(* IEC 61131-3 sources: Industry-PLC-LLM/data/PLCBEAD_repo/PLCBEAD_PLCEmbed-main/PLC-BEAD/Source/PLC_Programs (part 2) *)

(* ---- ALARM_2.ST ---- *)
FUNCTION_BLOCK ALARM_2
	VAR_INPUT
		X :	REAL;
		LO_1 :	REAL;
		HI_1 :	REAL;
		LO_2 :	REAL;
		HI_2 :	REAL;
		HYS :	REAL;
	END_VAR

	VAR_OUTPUT
		Q1_LO :	BOOL;
		Q1_HI :	BOOL;
		Q2_LO :	BOOL;
		Q2_HI :	BOOL;
	END_VAR

	VAR
		tmp :	REAL;
	END_VAR

	tmp := X - Hys * 0.5;
	IF tmp > LO_1 THEN Q1_LO := FALSE; END_IF;
	IF tmp > LO_2 THEN Q2_LO := FALSE; END_IF;
	IF tmp > HI_1 THEN Q1_HI := TRUE; END_IF;
	IF tmp > HI_2 THEN Q2_HI := TRUE; END_IF;
	tmp := tmp + hys;
	IF tmp < LO_1 THEN Q1_LO := TRUE; END_IF;
	IF tmp < LO_2 THEN Q2_LO := TRUE; END_IF;
	IF tmp < HI_1 THEN Q1_HI := FALSE; END_IF;
	IF tmp < HI_2 THEN Q2_HI := FALSE; END_IF;

END_FUNCTION_BLOCK

PROGRAM program0
	VAR
	    LocalVar0 : REAL;
		LocalVar1 : REAL;
		LocalVar2 : REAL;
		LocalVar3 : REAL;
		LocalVar4 : REAL;
		LocalVar5 : REAL;
		LocalOUT1  : BOOL;
		LocalOUT2  : BOOL;
		LocalOUT3  : BOOL;
		LocalOUT4  : BOOL;
		func_block : ALARM_2;
  	END_VAR
	func_block.X := LocalVar0;
	func_block.LO_1 := LocalVar1;
	func_block.HI_1 := LocalVar2;
	func_block.LO_2 := LocalVar3;
	func_block.HI_2 := LocalVar4;
	func_block.HYS := LocalVar5;
	func_block();
	LocalOUT1 := func_block.Q1_LO;
	LocalOUT2 := func_block.Q1_HI;
	LocalOUT3 := func_block.Q2_LO;
	LocalOUT4 := func_block.Q2_HI;
END_PROGRAM

CONFIGURATION Config0
  	RESOURCE Res0 ON PLC
    	TASK task0(INTERVAL := T#20ms,PRIORITY := 0);
    	PROGRAM instance0 WITH task0 : program0;
  	END_RESOURCE
END_CONFIGURATION

(* ---- ARRAY_AVG.ST ---- *)
TYPE
	oscat_pt_ARRAY: ARRAY [1..100] OF REAL;
END_TYPE

FUNCTION_BLOCK ARRAY_AVG_Block
	VAR_IN_OUT
		PT :	oscat_pt_ARRAY;
	END_VAR

	VAR_INPUT
		SIZE :	UINT;
	END_VAR

	VAR_OUTPUT
		ARRAY_AVG :	REAL;
	END_VAR

	VAR
		i :	INT;
		stop :	INT;
	END_VAR

	stop :=LIMIT_INT(1,UINT_TO_INT(size),1000);

	array_avg := 0.0;
	FOR i := 1 TO stop DO
		array_avg := array_avg + pt[i];
	END_FOR;
	array_avg := array_avg / INT_TO_REAL(stop);
END_FUNCTION_BLOCK

PROGRAM program0
  VAR
    LocalVar0 : oscat_pt_ARRAY;
    LocalVar1 : UINT;
	LocalOUT  : REAL;
	func_block : ARRAY_AVG_Block;
  END_VAR
	func_block.pt := LocalVar0;
	func_block.size := LocalVar1;
	func_block();
	LocalOUT := func_block.ARRAY_AVG;

END_PROGRAM

CONFIGURATION Config0
  RESOURCE Res0 ON PLC
    TASK task0(INTERVAL := T#20ms,PRIORITY := 0);
    PROGRAM instance0 WITH task0 : program0;
  END_RESOURCE
END_CONFIGURATION

(* ---- ARRAY_GAV.ST ---- *)
TYPE
	oscat_pt_ARRAY: ARRAY [1..100] OF REAL;
END_TYPE

FUNCTION SQRTN:REAL
	VAR_INPUT
		X :	REAL;
		N :	INT;
	END_VAR

	IF N > 0 THEN
		SQRTN := EXP(LN(x) / INT_TO_REAL(n));
	ELSE
		SQRTN := 0.0;
	END_IF;
END_FUNCTION

FUNCTION_BLOCK ARRAY_GAV_Block
	VAR_IN_OUT
		PT :	oscat_pt_ARRAY;
	END_VAR

	VAR_INPUT
		SIZE :	UINT;
	END_VAR

	VAR_OUTPUT
		ARRAY_GAV :	REAL;
	END_VAR

	VAR
		i :	INT;
		stop :	INT;
	END_VAR

	stop :=LIMIT_INT(1,UINT_TO_INT(size),1000);
	ARRAY_GAV := 1.0;
	FOR i := 1 TO stop DO
		IF pt[i] > 0.0 THEN
			ARRAY_GAV := ARRAY_GAV * pt[i];
		ELSE
			ARRAY_GAV := 0.0;
			RETURN;
		END_IF;
	END_FOR;
	ARRAY_GAV := SQRTN(ARRAY_GAV,stop);
END_FUNCTION_BLOCK

PROGRAM program0
  VAR
    LocalVar0 : oscat_pt_ARRAY;
    LocalVar1 : UINT;
	LocalOUT  : REAL;
	func_block : ARRAY_GAV_Block;
  END_VAR
	func_block.pt := LocalVar0;
	func_block.size := LocalVar1;
	func_block();
	LocalOUT := func_block.ARRAY_GAV;

END_PROGRAM

CONFIGURATION Config0
  RESOURCE Res0 ON PLC
    TASK task0(INTERVAL := T#20ms,PRIORITY := 0);
    PROGRAM instance0 WITH task0 : program0;
  END_RESOURCE
END_CONFIGURATION

(* ---- ARRAY_HAV.ST ---- *)
TYPE
	oscat_pt_ARRAY: ARRAY [1..100] OF REAL;
END_TYPE

FUNCTION_BLOCK ARRAY_HAV_Block
	VAR_IN_OUT
		PT :	oscat_pt_ARRAY;
	END_VAR

	VAR_INPUT
		SIZE :	UINT;
	END_VAR

	VAR_OUTPUT
		ARRAY_HAV :	REAL;
	END_VAR

	VAR
		i :	INT;
		stop :	INT;
	END_VAR

	stop :=LIMIT_INT(1,UINT_TO_INT(size),1000);
	ARRAY_HAV := 0.0;
	FOR i := 1 TO stop DO
		IF pt[i] <> 0.0 THEN
			ARRAY_HAV := ARRAY_HAV + 1.0/pt[i];
		ELSE
			ARRAY_HAV := 0.0;
			RETURN;
		END_IF;
	END_FOR;
	ARRAY_HAV := INT_TO_REAL(stop) / ARRAY_HAV;
END_FUNCTION_BLOCK

PROGRAM program0
  VAR
    LocalVar0 : oscat_pt_ARRAY;
    LocalVar1 : UINT;
	LocalOUT  : REAL;
	func_block : ARRAY_HAV_Block;
  END_VAR
	func_block.pt := LocalVar0;
	func_block.size := LocalVar1;
	func_block();
	LocalOUT := func_block.ARRAY_HAV;

END_PROGRAM

CONFIGURATION Config0
  RESOURCE Res0 ON PLC
    TASK task0(INTERVAL := T#20ms,PRIORITY := 0);
    PROGRAM instance0 WITH task0 : program0;
  END_RESOURCE
END_CONFIGURATION

(* ---- ARRAY_MAX.ST ---- *)
TYPE
	oscat_pt_ARRAY: ARRAY [1..100] OF REAL;
END_TYPE

FUNCTION_BLOCK ARRAY_MAX_Block
	VAR_IN_OUT
		PT :	oscat_pt_ARRAY;
	END_VAR

	VAR_INPUT
		SIZE :	UINT;
	END_VAR

	VAR_OUTPUT
		ARRAY_MAX :	REAL;
	END_VAR

	VAR
		i :	INT;
		stop :	INT;
	END_VAR

	stop :=LIMIT_INT(1,UINT_TO_INT(size),1000);

	FOR i := 1 TO stop DO
		IF pt[i] > array_max THEN array_max := pt[i]; END_IF;
	END_FOR;

END_FUNCTION_BLOCK

PROGRAM program0
  VAR
    LocalVar0 : oscat_pt_ARRAY;
    LocalVar1 : UINT;
	LocalOUT  : REAL;
	func_block : ARRAY_MAX_Block;
  END_VAR
	func_block.pt := LocalVar0;
	func_block.size := LocalVar1;
	func_block();
	LocalOUT := func_block.ARRAY_MAX;

END_PROGRAM

CONFIGURATION Config0
  RESOURCE Res0 ON PLC
    TASK task0(INTERVAL := T#20ms,PRIORITY := 0);
    PROGRAM instance0 WITH task0 : program0;
  END_RESOURCE
END_CONFIGURATION

(* ---- ARRAY_MEDIAN.ST ---- *)
TYPE
	oscat_pt_ARRAY: ARRAY [1..100] OF REAL;
	oscat_stack_array: ARRAY [1..32]   OF INT;
END_TYPE

FUNCTION _INT_TO_UDINT:UDINT
	VAR_INPUT
		IN :	INT;
	END_VAR

	_INT_TO_UDINT := DINT_TO_UDINT(INT_TO_DINT(IN));
END_FUNCTION

FUNCTION BIT_OF_DWORD:BOOL
	VAR_INPUT
		IN :	DWORD;
		N :	INT;
	END_VAR
	BIT_OF_DWORD := (SHR(in,n) AND DWORD#1) > DWORD#0;
END_FUNCTION

FUNCTION EVEN:BOOL
	VAR_INPUT
		IN :	DINT;
	END_VAR
	even := NOT BIT_OF_DWORD(DINT_TO_DWORD(in),0);
END_FUNCTION

FUNCTION_BLOCK _ARRAY_SORT_Block
	VAR_IN_OUT
		PT :	oscat_pt_ARRAY;
	END_VAR

	VAR_INPUT
		SIZE :	UINT;
	END_VAR

	VAR_OUTPUT
		_ARRAY_SORT :BOOL;
	END_VAR

	VAR
		stack_count :	INT;
		stack :	oscat_stack_array;
		links :	INT;
		rechts :	INT;
		pivot :	REAL;
		i :	INT;
		j :	INT;
		ende_innen :	BOOL;
		ende_aussen :	BOOL;
		tmp :	REAL;
		x :	INT;
	END_VAR

	links := 1;
	rechts := DWORD_TO_INT(SHR(UINT_TO_DWORD(size),2));
	stack_count := 1;

	WHILE NOT ende_aussen DO
		IF links < rechts THEN
			x := DWORD_TO_INT(SHR(UDINT_TO_DWORD(_INT_TO_UDINT(rechts)+ _INT_TO_UDINT(links)),1));
			pivot := PT[x];
			i := links - 1;
			j := rechts + 1;

			ende_innen := FALSE;
			REPEAT
				REPEAT	i := i+1;	UNTIL (PT[i] >= pivot) OR NOT (i < rechts)	END_REPEAT;
				REPEAT	j := j-1;	UNTIL (PT[j] <= pivot) OR NOT (j > links)	END_REPEAT;
				IF i >= j THEN
					ende_innen := TRUE;
				ELSE
					tmp := PT[j];
					PT[j] := PT[i];
					PT[i] := tmp;
				END_IF;

			UNTIL ende_innen END_REPEAT;

			stack[stack_count] := rechts;
			IF Stack_count < 32 THEN
				stack_count := stack_count +1;
			ELSE
				ende_aussen := TRUE;
				_ARRAY_SORT := FALSE;
			END_IF;
			rechts := MAX(links, i-1);

		ELSE
			IF stack_count = 1 THEN
				ende_aussen := TRUE;
			ELSE
				links := rechts+1;
				stack_count := stack_count - 1;
				rechts:= stack[stack_count];
			END_IF;
		END_IF;
	END_WHILE;

	_ARRAY_SORT := TRUE;
END_FUNCTION_BLOCK

FUNCTION_BLOCK _ARRAY_MEDIAN_Block

	VAR_IN_OUT
		PT :	oscat_pt_ARRAY;
	END_VAR

	VAR_INPUT
		SIZE :	UINT;
	END_VAR

	VAR_OUTPUT
		_ARRAY_MEDIAN :	REAL;
	END_VAR

	VAR
		i :	INT;
		i2 :	INT;
		stop :	INT;
		_array_sort :	_ARRAY_SORT_Block;
	END_VAR

	(* Array sortieren *)
	_array_sort.pt   := pt;
	_array_sort.size := size;
	_array_sort();
	pt := _array_sort.pt;

	stop :=LIMIT_INT(1,UINT_TO_INT(size),1000);
	IF even(INT_TO_DINT(stop)) THEN
	    i := WORD_TO_INT(SHR(INT_TO_WORD(stop),1));
	    i2 := i+1;
		_array_median := (pt[i] + pt[i2]) * 0.5;
	ELSE
	    i := WORD_TO_INT(SHR(INT_TO_WORD(stop),1))+1;
		_array_median := pt[i];
	END_IF;

END_FUNCTION_BLOCK

PROGRAM program0
  VAR
    LocalVar0 : oscat_pt_ARRAY;
    LocalVar1 : UINT;
	LocalOUT  : REAL;
	func_block : _ARRAY_MEDIAN_Block;
  END_VAR
	func_block.pt := LocalVar0;
	func_block.size := LocalVar1;
	func_block();
	LocalOUT := func_block._ARRAY_MEDIAN;
	LocalVar0 := func_block.pt;

END_PROGRAM

CONFIGURATION Config0
  RESOURCE Res0 ON PLC
    TASK task0(INTERVAL := T#20ms,PRIORITY := 0);
    PROGRAM instance0 WITH task0 : program0;
  END_RESOURCE
END_CONFIGURATION

(* ---- ARRAY_MIN.ST ---- *)
TYPE
	oscat_pt_ARRAY: ARRAY [1..100] OF REAL;
END_TYPE

FUNCTION_BLOCK ARRAY_MIN_Block
	VAR_IN_OUT
		PT :	oscat_pt_ARRAY;
	END_VAR

	VAR_INPUT
		SIZE :	UINT;
	END_VAR

	VAR_OUTPUT
		ARRAY_MIN :	REAL;
	END_VAR

	VAR
		i :	INT;
		stop :	INT;
	END_VAR

	stop :=LIMIT_INT(1,UINT_TO_INT(size),1000);

	array_min := pt[1];
	FOR i := 2 TO stop DO
		IF pt[i] < array_min THEN array_min := pt[i]; END_IF;
	END_FOR;

END_FUNCTION_BLOCK
PROGRAM program0
  VAR
    LocalVar0 : oscat_pt_ARRAY;
    LocalVar1 : UINT;
	LocalOUT  : REAL;
	func_block : ARRAY_MIN_Block;
  END_VAR
	func_block.pt := LocalVar0;
	func_block.size := LocalVar1;
	func_block();
	LocalOUT := func_block.ARRAY_MIN;

END_PROGRAM

CONFIGURATION Config0
  RESOURCE Res0 ON PLC
    TASK task0(INTERVAL := T#20ms,PRIORITY := 0);
    PROGRAM instance0 WITH task0 : program0;
  END_RESOURCE
END_CONFIGURATION

(* ---- ARRAY_SDV.ST ---- *)
TYPE
	oscat_pt_ARRAY: ARRAY [1..100] OF REAL;
END_TYPE

FUNCTION_BLOCK ARRAY_VAR_Block
	VAR_IN_OUT
		PT :	oscat_pt_ARRAY;
	END_VAR

	VAR_INPUT
		SIZE :	UINT;
	END_VAR

	VAR_OUTPUT
		ARRAY_VAR :	REAL;
	END_VAR

	VAR
		i :	INT;
		stop :	INT;
		avg :	REAL;
	END_VAR

	stop :=LIMIT_INT(1,UINT_TO_INT(size),1000);
	avg := pt[1];
	FOR i := 2 TO stop DO
		avg := avg + pt[i];
	END_FOR;
	avg := avg / INT_TO_REAL(stop);

	array_var := EXPT(pt[1] - avg, 2.0);
	FOR i := 2 TO stop DO
		array_var := array_var + EXPT(pt[i] - avg, 2.0);
	END_FOR;
	array_var := array_var / INT_TO_REAL(stop-1);

END_FUNCTION_BLOCK

FUNCTION_BLOCK ARRAY_SDV_Block
	VAR_IN_OUT
		PT :	oscat_pt_ARRAY;
	END_VAR

	VAR_INPUT
		SIZE :	UINT;
	END_VAR

	VAR_OUTPUT
		ARRAY_SDV :	REAL;
	END_VAR

	VAR
		FB_array_var :	array_var_block;
	END_VAR

	FB_array_var.pt   := pt;
	FB_array_var.size := size;
	FB_array_var();
	pt := FB_array_var.pt;

	array_sdv := SQRT(FB_array_var.array_var);
END_FUNCTION_BLOCK

PROGRAM program0
  VAR
    LocalVar0 : oscat_pt_ARRAY;
    LocalVar1 : UINT;
	LocalOUT  : REAL;
	func_block : ARRAY_SDV_Block;
  END_VAR
	func_block.pt := LocalVar0;
	func_block.size := LocalVar1;
	func_block();
	LocalOUT := func_block.ARRAY_SDV;

END_PROGRAM

CONFIGURATION Config0
  RESOURCE Res0 ON PLC
    TASK task0(INTERVAL := T#20ms,PRIORITY := 0);
    PROGRAM instance0 WITH task0 : program0;
  END_RESOURCE
END_CONFIGURATION

(* ---- ARRAY_SPR.ST ---- *)
TYPE
	oscat_pt_ARRAY: ARRAY [1..100] OF REAL;
END_TYPE

FUNCTION_BLOCK ARRAY_SPR_Block
	VAR_IN_OUT
		PT :	oscat_pt_ARRAY;
	END_VAR

	VAR_INPUT
		SIZE :	UINT;
	END_VAR

	VAR_OUTPUT
		ARRAY_SPR :	REAL;
	END_VAR

	VAR
		i :	INT;
		stop :	INT;
		array_max :	REAL;
		array_min :	REAL;
	END_VAR

	stop :=LIMIT_INT(1,UINT_TO_INT(size),1000);

	array_min := pt[1];
	array_max := pt[1];
	FOR i := 2 TO stop DO
		IF pt[i] > array_max THEN array_max := pt[i];
		ELSIF pt[i] < array_min THEN array_min := pt[i];
		END_IF;
	END_FOR;
	array_spr := array_max - array_min;
END_FUNCTION_BLOCK

PROGRAM program0
  VAR
    LocalVar0 : oscat_pt_ARRAY;
    LocalVar1 : UINT;
	LocalOUT  : REAL;
	func_block : ARRAY_SPR_Block;
  END_VAR
	func_block.pt := LocalVar0;
	func_block.size := LocalVar1;
	func_block();
	LocalOUT := func_block.ARRAY_SPR;

END_PROGRAM

CONFIGURATION Config0
  RESOURCE Res0 ON PLC
    TASK task0(INTERVAL := T#20ms,PRIORITY := 0);
    PROGRAM instance0 WITH task0 : program0;
  END_RESOURCE
END_CONFIGURATION

(* ---- ARRAY_SUM.ST ---- *)
TYPE
	oscat_pt_ARRAY: ARRAY [1..100] OF REAL;
END_TYPE

FUNCTION_BLOCK ARRAY_SUM_Block
	VAR_IN_OUT
		PT :	oscat_pt_ARRAY;
	END_VAR

	VAR_INPUT
		SIZE :	UINT;
	END_VAR

	VAR_OUTPUT
		ARRAY_SUM :	REAL;
	END_VAR

	VAR
		i :	INT;
		stop :	INT;
	END_VAR

	stop :=LIMIT_INT(1,UINT_TO_INT(size),1000);

	array_sum := pt[1];
	FOR i := 2 TO stop DO
		array_sum := array_sum + pt[i];
	END_FOR;
END_FUNCTION_BLOCK

PROGRAM program0
  VAR
    LocalVar0 : oscat_pt_ARRAY;
    LocalVar1 : UINT;
	LocalOUT  : REAL;
	func_block : ARRAY_SUM_Block;
  END_VAR
	func_block.pt := LocalVar0;
	func_block.size := LocalVar1;
	func_block();
	LocalOUT := func_block.ARRAY_SUM;

END_PROGRAM

CONFIGURATION Config0
  RESOURCE Res0 ON PLC
    TASK task0(INTERVAL := T#20ms,PRIORITY := 0);
    PROGRAM instance0 WITH task0 : program0;
  END_RESOURCE
END_CONFIGURATION

(* ---- ARRAY_TREND.ST ---- *)
TYPE
	oscat_pt_ARRAY: ARRAY [1..100] OF REAL;
END_TYPE

FUNCTION BIT_OF_DWORD:BOOL
	VAR_INPUT
		IN :	DWORD;
		N :	INT;
	END_VAR
	BIT_OF_DWORD := (SHR(in,n) AND DWORD#1) > DWORD#0;
END_FUNCTION

FUNCTION EVEN:BOOL
	VAR_INPUT
		IN :	DINT;
	END_VAR
	even := NOT BIT_OF_DWORD(DINT_TO_DWORD(in),0);
END_FUNCTION

FUNCTION_BLOCK ARRAY_TREND_Block
	VAR_IN_OUT
		PT :	oscat_pt_ARRAY;
	END_VAR

	VAR_INPUT
		SIZE :	UINT;
	END_VAR

	VAR_OUTPUT
		ARRAY_TREND :	REAL;
	END_VAR

	VAR
		d :	INT;
		i :	INT;
		stop :	INT;
		stop2 :	INT;
		x :	REAL;
	END_VAR

	x := 0.0;
	stop :=LIMIT_INT(1,UINT_TO_INT(size),1000);
	stop2 := WORD_TO_INT(SHR(INT_TO_WORD(stop),1));
	IF even(INT_TO_DINT(stop)) THEN d:=0; ELSE d:=1;END_IF;

	FOR i := 1 TO stop2+d DO
		x := x - pt[i];
	END_FOR;
	FOR i := stop2+1 TO stop DO
		x := x + pt[i];
	END_FOR;
	array_trend := x / INT_TO_REAL(stop2+d);

END_FUNCTION_BLOCK

PROGRAM program0
  VAR
    LocalVar0 : oscat_pt_ARRAY;
    LocalVar1 : UINT;
	LocalOUT  : REAL;
	func_block : ARRAY_TREND_Block;
  END_VAR
	func_block.pt := LocalVar0;
	func_block.size := LocalVar1;
	func_block();
	LocalOUT := func_block.ARRAY_TREND;

END_PROGRAM

CONFIGURATION Config0
  RESOURCE Res0 ON PLC
    TASK task0(INTERVAL := T#20ms,PRIORITY := 0);
    PROGRAM instance0 WITH task0 : program0;
  END_RESOURCE
END_CONFIGURATION

(* ---- ARRAY_VAR.ST ---- *)
TYPE
	oscat_pt_ARRAY: ARRAY [1..100] OF REAL;
END_TYPE

FUNCTION_BLOCK ARRAY_VAR_Block
	VAR_IN_OUT
		PT :	oscat_pt_ARRAY;
	END_VAR

	VAR_INPUT
		SIZE :	UINT;
	END_VAR

	VAR_OUTPUT
		ARRAY_VAR :	REAL;
	END_VAR

	VAR
		i :	INT;
		stop :	INT;
		avg :	REAL;
	END_VAR

	stop :=LIMIT_INT(1,UINT_TO_INT(size),1000);
	avg := pt[1];
	FOR i := 2 TO stop DO
		avg := avg + pt[i];
	END_FOR;
	avg := avg / INT_TO_REAL(stop);

	array_var := EXPT(pt[1] - avg, 2.0);
	FOR i := 2 TO stop DO
		array_var := array_var + EXPT(pt[i] - avg, 2.0);
	END_FOR;
	array_var := array_var / INT_TO_REAL(stop-1);

END_FUNCTION_BLOCK

PROGRAM program0
  VAR
    LocalVar0 : oscat_pt_ARRAY;
    LocalVar1 : UINT;
	LocalOUT  : REAL;
	func_block : ARRAY_VAR_Block;
  END_VAR
	func_block.pt := LocalVar0;
	func_block.size := LocalVar1;
	func_block();
	LocalOUT := func_block.ARRAY_VAR;

END_PROGRAM

CONFIGURATION Config0
  RESOURCE Res0 ON PLC
    TASK task0(INTERVAL := T#20ms,PRIORITY := 0);
    PROGRAM instance0 WITH task0 : program0;
  END_RESOURCE
END_CONFIGURATION

(* ---- ASTRO.ST ---- *)
FUNCTION_BLOCK ASTRO
	VAR_INPUT
		M :	REAL;
		AE :	REAL;
		PC :	REAL;
		LJ :	REAL;
	END_VAR

	VAR_OUTPUT
		YM :	REAL;
		YAE :	REAL;
		YPC :	REAL;
		YLJ :	REAL;
	END_VAR

	YAE :=	AE
			+ m * 6.6845871535E-012
			+ PC * 206265.0
			+ LJ * 63240.0;
	Ym := YAE * 149.597870E9;
	YPC := YAE * 4.8481322570E-006;
	YLJ := YAE * 1.5812776724E-005;
END_FUNCTION_BLOCK

PROGRAM program0
  VAR
    LocalVar0 : REAL;
    LocalVar1 : REAL;
	LocalVar2 : REAL;
	LocalVar3 : REAL;
	LocalOUT1 : REAL;
	LocalOUT2 : REAL;
	LocalOUT3 : REAL;
	LocalOUT4 : REAL;
	func_block : ASTRO;
  END_VAR
	func_block.M  := LocalVar0;
	func_block.AE := LocalVar1;
	func_block.PC := LocalVar2;
	func_block.LJ := LocalVar3;
	func_block();
	LocalOUT1 := func_block.YM ;
	LocalOUT2 := func_block.YAE;
	LocalOUT3 := func_block.YPC;
	LocalOUT4 := func_block.YLJ;

END_PROGRAM

CONFIGURATION Config0
  RESOURCE Res0 ON PLC
    TASK task0(INTERVAL := T#20ms,PRIORITY := 0);
    PROGRAM instance0 WITH task0 : program0;
  END_RESOURCE
END_CONFIGURATION

(* ---- AUTORUN.ST ---- *)
FUNCTION UDINT_TO_TIME2:TIME

	VAR_INPUT
		IN :	UDINT;
	END_VAR

	UDINT_TO_TIME2 := DINT_TO_TIME(UDINT_TO_DINT(IN));

END_FUNCTION

FUNCTION_BLOCK T_PLC_MS_block
	VAR_OUTPUT
		T_PLC_MS :	UDINT;
	END_VAR

	VAR_EXTERNAL
		PLC_TICKS_PER_SEC :	INT;
		PLC_SYS_TICK_CNT :	DINT;
	END_VAR

	VAR
		debug :	BOOL;(*Debug-Mode ON / OFF*)
		N :	INT;(*Debug-Faktor*)
		Offset :	UDINT;(*Debug-Offset*)
		temp :	DWORD := DWORD#1;(*Debug-Offset*)
		mode :	BOOL;(*modus*)
		faktor :	UDINT;(*Systemtakt-Faktor*)
		init :	BOOL;
		v_plc_ticks_per_sec :	UDINT;
		base :	UDINT := UDINT#1000;
	END_VAR

	IF init = FALSE THEN
		v_plc_ticks_per_sec := INT_TO_UDINT(PLC_TICKS_PER_SEC);
		IF v_plc_ticks_per_sec = UDINT#1024 THEN
			faktor := UDINT#1;
			mode := FALSE;
		ELSIF v_plc_ticks_per_sec > UDINT#0 THEN
			IF v_plc_ticks_per_sec <= base THEN
				faktor := base / v_plc_ticks_per_sec;
				mode := FALSE;
			ELSE
				faktor := v_plc_ticks_per_sec / base;
				mode := TRUE;
			END_IF;
		ELSE
			faktor := UDINT#1;
		END_IF;
		init := TRUE;
	END_IF;

	IF mode THEN
		T_PLC_MS := DINT_TO_UDINT(PLC_SYS_TICK_CNT) / faktor;
	ELSE
		T_PLC_MS := DINT_TO_UDINT(PLC_SYS_TICK_CNT) * faktor;
	END_IF;

	IF debug THEN
		T_PLC_MS := (DWORD_TO_UDINT(SHL(UDINT_TO_DWORD(T_PLC_MS),N) OR SHL(temp,N)) - UDINT#1) + Offset;
	END_IF;

END_FUNCTION_BLOCK

FUNCTION TIME_TO_UDINT2:UDINT
	VAR_INPUT
		X :	TIME;
	END_VAR

	TIME_TO_UDINT2 := DINT_TO_UDINT(TIME_TO_DINT(X));
END_FUNCTION

FUNCTION FRMP_B:BYTE
	VAR_INPUT
		START :	BYTE;
		DIR :	BOOL;
		TD :	TIME;
		TR :	TIME;
	END_VAR

	IF TD < TR THEN
		FRMP_B := MIN(UDINT_TO_BYTE(DWORD_TO_UDINT(SHL(TIME_TO_DWORD(TD), 8)) / TIME_TO_UDINT2(TR)), SEL(DIR, START, USINT_TO_BYTE(USINT#255 - BYTE_TO_USINT(START))));
		IF DIR THEN
			FRMP_B := USINT_TO_BYTE(BYTE_TO_USINT(START) + BYTE_TO_USINT(FRMP_B));
		ELSE
			FRMP_B := USINT_TO_BYTE(BYTE_TO_USINT(START) - BYTE_TO_USINT(FRMP_B));
		END_IF;
	ELSE
		FRMP_B := SEL(DIR, BYTE#0, BYTE#255);
	END_IF;
END_FUNCTION

FUNCTION_BLOCK _RMP_B
	VAR_INPUT
		DIR :	BOOL;
		E :	BOOL := TRUE;
		TR :	TIME;
	END_VAR

	VAR_IN_OUT
		RMP :	BYTE;
	END_VAR

	VAR
		T_PLC_MS :	T_PLC_MS_block;
		tx :	TIME;
		tl :	TIME;
		tn :	TIME;
		init :	BOOL;
		last_dir :	BOOL;
		start :	BYTE;
	END_VAR

	T_PLC_MS();
	tx := UDINT_TO_TIME(T_PLC_MS.T_PLC_MS);

	IF E AND init AND (dir = last_dir) AND (RMP <> SEL(DIR, BYTE#0, BYTE#255)) AND TR = tn THEN
		RMP := FRMP_B(start, DIR, tx - tl, TR);
	ELSE
		init := TRUE;
		tl := tx;
		tn := tr;
		start := RMP;
	END_IF;
	last_dir := dir;
END_FUNCTION_BLOCK

FUNCTION_BLOCK AUTORUN_Block

	VAR_INPUT
		IN :	BOOL;
		TEST :	BOOL;
		ARE :	BOOL := TRUE;
		TRUN :	TIME;
		TOFF :	TIME;
	END_VAR

	VAR_OUTPUT
		OUT :	BOOL;
		ARO :	BOOL;
	END_VAR

	VAR_IN_OUT
		ARX :	BOOL;
	END_VAR

	VAR
		timer :	_RMP_B;
		val :	BYTE;
	END_VAR

	IF TOFF > T#0s THEN
		timer(DIR:= OUT, TR := SEL(OUT, TOFF, TRUN), RMP := val);
		val := timer.RMP;
	ELSE
		val := BYTE#255;
	END_IF;

	IF (NOT ARX AND ARE AND val = BYTE#0) OR TEST THEN
		val := BYTE#0;
		ARO := TRUE;
		ARX := TRUE;
	ELSIF val = BYTE#255 AND ARO THEN
		ARO := FALSE;
		ARX := FALSE;
	END_IF;

	out := IN OR ARO;

END_FUNCTION_BLOCK

PROGRAM program0
	VAR
		IN :	BOOL;
		TEST :	BOOL;
		ARE :	BOOL := TRUE;
		TRUN :	TIME;
		TOFF :	TIME;
		OUT :	BOOL;
		ARO :	BOOL;
		func_block : AUTORUN_Block;
	END_VAR
	func_block.IN := IN;
	func_block.TEST := TEST;
	func_block.ARE := ARE ;
	func_block.TRUN := TRUN;
	func_block.TOFF := TOFF;
	func_block();
	OUT  := func_block.OUT;
	ARO  := func_block.ARO;
END_PROGRAM

CONFIGURATION Config0
	VAR_GLOBAL
		PLC_TICKS_PER_SEC :	INT;
		PLC_SYS_TICK_CNT :	DINT;
	END_VAR
  	RESOURCE Res0 ON PLC
    	TASK task0(INTERVAL := T#20ms,PRIORITY := 0);
    	PROGRAM instance0 WITH task0 : program0;
  	END_RESOURCE
END_CONFIGURATION

(* ---- B_TRIG.ST ---- *)
FUNCTION_BLOCK B_TRIG
	VAR_INPUT
		CLK :	BOOL;
	END_VAR

	VAR_OUTPUT
		Q :	BOOL := FALSE;
	END_VAR

	VAR
		edge :	BOOL := FALSE;
	END_VAR

	Q := clk XOR edge;
	edge := CLK;
END_FUNCTION_BLOCK

PROGRAM program0
  VAR
    LocalVar0 : BOOL;
	LocalOUT  : BOOL;
	func_block : B_TRIG;
  END_VAR
	func_block.CLK := LocalVar0;
	func_block();
	LocalOUT := func_block.Q;

END_PROGRAM

CONFIGURATION Config0
  RESOURCE Res0 ON PLC
    TASK task0(INTERVAL := T#20ms,PRIORITY := 0);
    PROGRAM instance0 WITH task0 : program0;
  END_RESOURCE
END_CONFIGURATION

(* ---- BAR_GRAPH.ST ---- *)
FUNCTION_BLOCK BAR_GRAPH
	VAR_INPUT
		X :	REAL;
		RST :	BOOL;
		TRIGGER_LOW :	REAL;
		TRIGGER_HIGH :	REAL;
		ALARM_LOW :	BOOL;
		ALARM_HIGH :	BOOL;
		LOG_SCALE :	BOOL;
	END_VAR

	VAR_OUTPUT
		LOW :	BOOL;
		Q1 :	BOOL;
		Q2 :	BOOL;
		Q3 :	BOOL;
		Q4 :	BOOL;
		Q5 :	BOOL;
		Q6 :	BOOL;
		HIGH :	BOOL;
		ALARM :	BOOL;
		STATUS :	BYTE;
	END_VAR

	VAR
		init :	BOOL;
		T1 :	REAL;
		T2 :	REAL;
		T3 :	REAL;
		T4 :	REAL;
		T5 :	REAL;
		temp :	REAL;
	END_VAR

	IF NOT init THEN
		init := TRUE;
		IF log_scale THEN
			temp := EXP(LN(Trigger_high / Trigger_low) * 0.166666666666666666666);
			T1 := trigger_low * temp;
			T2 := T1 * temp;
			T3 := T2 * temp;
			T4 := T3 * temp;
			T5 := T4 * temp;
		ELSE
			temp := (trigger_high - trigger_low) * 0.142857142;
			T1 := trigger_low + temp;
			T2 := T1 + temp;
			T3 := T2 + temp;
			T4 := T3 + temp;
			T5 := T4 + temp;
		END_IF;
	END_IF;

	Q1 := FALSE;
	Q2 := FALSE;
	Q3 := FALSE;
	Q4 := FALSE;
	Q5 := FALSE;
	Q6 := FALSE;
	status := BYTE#110;

	IF NOT alarm_low THEN low := FALSE; END_IF;
	IF NOT alarm_high THEN high := FALSE; END_IF;
	IF rst THEN
		alarm := FALSE;
		low := FALSE;
		high := FALSE;
	END_IF;

	IF X < trigger_low THEN
		Low := TRUE;
		status := BYTE#111;
		IF alarm_low THEN
			alarm := TRUE;
			status := BYTE#1;
		END_IF;
	ELSIF X < T1 THEN
		Q1 := TRUE;
	ELSIF x < t2 THEN
		Q2 := TRUE;
	ELSIF x < t3 THEN
		Q3 := TRUE;
	ELSIF x < T4 THEN
		Q4 := TRUE;
	ELSIF x < T5 THEN
		q5 := TRUE;
	ELSIF x < trigger_high THEN
		q6 := TRUE;
	ELSE
		high := TRUE;
		status := BYTE#112;
		IF alarm_high THEN
			alarm := TRUE;
			status := BYTE#2;
		END_IF;
	END_IF;

END_FUNCTION_BLOCK

PROGRAM program0
  VAR
    LocalVar0 : REAL;
    LocalVar1 : BOOL;
	LocalVar2 : REAL;
	LocalVar3 : REAL;
	LocalVar4 : BOOL;
	LocalVar5 : BOOL;
	LocalVar6 : BOOL;

	LOW   :	BOOL;
	Q1    :	BOOL;
	Q2    :	BOOL;
	Q3    :	BOOL;
	Q4    :	BOOL;
	Q5    :	BOOL;
	Q6    :	BOOL;
	HIGH  :	BOOL;
	ALARM :	BOOL;
	STATUS:	BYTE;

	func_block : BAR_GRAPH;
  END_VAR
	func_block.X := LocalVar0;
	func_block.RST := LocalVar1;
	func_block.TRIGGER_LOW := LocalVar2;
	func_block.TRIGGER_HIGH := LocalVar3;
	func_block.ALARM_LOW := LocalVar4;
	func_block.ALARM_HIGH := LocalVar5;
	func_block.LOG_SCALE := LocalVar6;

	func_block();
	LOW   := func_block.LOW   ;
	Q1    := func_block.Q1    ;
	Q2    := func_block.Q2    ;
	Q3    := func_block.Q3    ;
	Q4    := func_block.Q4    ;
	Q5    := func_block.Q5    ;
	Q6    := func_block.Q6    ;
	HIGH  := func_block.HIGH  ;
	ALARM := func_block.ALARM ;
	STATUS:= func_block.STATUS;

END_PROGRAM

CONFIGURATION Config0
  RESOURCE Res0 ON PLC
    TASK task0(INTERVAL := T#20ms,PRIORITY := 0);
    PROGRAM instance0 WITH task0 : program0;
  END_RESOURCE
END_CONFIGURATION

(* ---- BASE64_DECODE_STR.ST ---- *)
TYPE
  oscat_aB0_47	: ARRAY [0..47]	OF BYTE;
  oscat_aB0_63	: ARRAY [0..63]	OF BYTE;
END_TYPE

FUNCTION_BLOCK BASE64_DECODE_STREAM
	VAR_IN_OUT
		BUF1 :	oscat_aB0_63;
		BUF2 :	oscat_aB0_47;
	END_VAR

	VAR_INPUT
		SIZE1 :	INT;
	END_VAR

	VAR_OUTPUT
		SIZE2 :	INT;
	END_VAR

	VAR
		a :	INT;
		b :	WORD;
		o :	INT;
		off :	INT;
		i1 :	INT;
		i2 :	INT;
		c :	INT;
	END_VAR

	IF SIZE1 <= 0 THEN SIZE2 := 0; RETURN; END_IF;
	c := SIZE1 - 1;
	i2 := 0;
	a := 0;
	b := WORD#0;
	FOR i1 := 0 TO c DO
		o := BYTE_TO_INT(BUF1[i1]);
		IF o = 61  (* = *) THEN EXIT;
		ELSIF o > 96 (* a-z *) THEN off := 71;
		ELSIF o > 64 (* A-Z *) THEN off := 65;
		ELSIF o > 47 (* 0-9 *) THEN off := -4;
		ELSIF o = 43 (* + *) THEN off := -19;
		ELSIF o = 47 (* / *) THEN off := -16;
		END_IF;
		b := SHL(b,6) OR INT_TO_WORD(o - off);
		a := a + 6;
		IF a >= 8 THEN
			a := a - 8;
			BUF2[i2] := WORD_TO_BYTE(SHR(b,a));
			i2 := i2 + 1;
			b := b AND NOT SHL(WORD#16#FFFF,a);
		END_IF;
	END_FOR;
	SIZE2 := i2;
END_FUNCTION_BLOCK

FUNCTION_BLOCK BASE64_DECODE_STR
	VAR_INPUT
		RUN :	BOOL;
	END_VAR

	VAR_OUTPUT
		DONE :	BOOL;
	END_VAR

	VAR_IN_OUT
		STR1 :	STRING;
		STR2 :	STRING;
	END_VAR

	VAR
		BASE64_DECODE_STREAM :	BASE64_DECODE_STREAM;
		run_last :	BOOL;
		buf1 :	oscat_aB0_63;
		buf2 :	oscat_aB0_47;
		mode :	INT;
		size1 :	INT;
		size2 :	INT;
		end :	INT;
		pos :	INT;
		i1 :	INT;
		i2 :	INT;
		i3 :	INT;
		STRx :	STRING;
		BTS :	BUF_TO_STRING;
	END_VAR

	(*@KEY@: WORKSHEET
	NAME: BASE64_DECODE_STR
	IEC_LANGUAGE: ST
	*)

	CASE mode OF
	0:	IF RUN AND NOT run_last THEN
			DONE := FALSE;
			mode := 1;
			end := LEN(STR1);
			pos := 0;
			STR2 := '';
		END_IF;
	1:
		SIZE1 := MIN(48,end - pos);
		IF SIZE1 > 0 THEN

			i2 := SIZE1 - 1;
			i3 := pos + 1;
			FOR i1 := 0 TO i2 DO
				buf1[i1] := INT_TO_BYTE(GET_CHAR(STR1,i3));
				i3 := i3 + 1;
			END_FOR;

			BASE64_DECODE_STREAM(BUF1:=BUF1 ,BUF2:=BUF2 ,SIZE1:=SIZE1);
			buf1  :=BASE64_DECODE_STREAM.BUF1;
			buf2  :=BASE64_DECODE_STREAM.BUF2;
			SIZE2 :=BASE64_DECODE_STREAM.SIZE2;

			FOR i1 := 0 TO 1 DO
				BTS.REQ := i1 > 0;
				BTS.BUF_FORMAT := TRUE;
				BTS.BUF_OFFS := DINT#0;
				BTS.BUF_CNT := INT_TO_DINT(SIZE2);
				BTS.BUFFER := buf2;
				BTS.DST := STRx;
				BTS();
				buf2 := BTS.BUFFER;
				STRx := BTS.DST;
			END_FOR;
			STR2 := CONCAT(STR2,STRx);
		ELSE
			mode := 0;
			DONE := TRUE;
		END_IF;
		pos := pos + size1;
	END_CASE;

	run_last := RUN;

END_FUNCTION_BLOCK

(* ---- BASE64_DECODE_STREAM.ST ---- *)
TYPE
  oscat_aB0_47	: ARRAY [0..47]	OF BYTE;
  oscat_aB0_63	: ARRAY [0..63]	OF BYTE;
END_TYPE

FUNCTION_BLOCK BASE64_DECODE_STREAM
	VAR_IN_OUT
		BUF1 :	oscat_aB0_63;
		BUF2 :	oscat_aB0_47;
	END_VAR

	VAR_INPUT
		SIZE1 :	INT;
	END_VAR

	VAR_OUTPUT
		SIZE2 :	INT;
	END_VAR

	VAR
		a :	INT;
		b :	WORD;
		o :	INT;
		off :	INT;
		i1 :	INT;
		i2 :	INT;
		c :	INT;
	END_VAR

	IF SIZE1 <= 0 THEN SIZE2 := 0; RETURN; END_IF;
	c := SIZE1 - 1;
	i2 := 0;
	a := 0;
	b := WORD#0;
	FOR i1 := 0 TO c DO
		o := BYTE_TO_INT(BUF1[i1]);
		IF o = 61  (* = *) THEN EXIT;
		ELSIF o > 96 (* a-z *) THEN off := 71;
		ELSIF o > 64 (* A-Z *) THEN off := 65;
		ELSIF o > 47 (* 0-9 *) THEN off := -4;
		ELSIF o = 43 (* + *) THEN off := -19;
		ELSIF o = 47 (* / *) THEN off := -16;
		END_IF;
		b := SHL(b,6) OR INT_TO_WORD(o - off);
		a := a + 6;
		IF a >= 8 THEN
			a := a - 8;
			BUF2[i2] := WORD_TO_BYTE(SHR(b,a));
			i2 := i2 + 1;
			b := b AND NOT SHL(WORD#16#FFFF,a);
		END_IF;
	END_FOR;
	SIZE2 := i2;
END_FUNCTION_BLOCK

PROGRAM program0
  VAR
	BUF1  :	oscat_aB0_63;
	BUF2  :	oscat_aB0_47;

	SIZE1 :	INT;

	SIZE2 :	INT;
	func_block : BASE64_DECODE_STREAM;
  END_VAR
	func_block.BUF1 :=BUF1 ;
	func_block.BUF2 :=BUF2 ;
	func_block.SIZE1:=SIZE1;
	func_block();
	BUF1 := func_block.BUF1;
	BUF2 := func_block.BUF2;
	SIZE2 := func_block.SIZE2;
END_PROGRAM

CONFIGURATION Config0
  RESOURCE Res0 ON PLC
    TASK task0(INTERVAL := T#20ms,PRIORITY := 0);
    PROGRAM instance0 WITH task0 : program0;
  END_RESOURCE
END_CONFIGURATION

(* ---- BASE64_ENCODE_STREAM.ST ---- *)
TYPE
  oscat_aB0_47	: ARRAY [0..47]	OF BYTE;
  oscat_aB0_63	: ARRAY [0..63]	OF BYTE;
END_TYPE

FUNCTION_BLOCK BASE64_ENCODE_STREAM

	VAR_IN_OUT
		BUF1 :	oscat_aB0_47;
		BUF2 :	oscat_aB0_63;
	END_VAR

	VAR_INPUT
		SIZE1 :	INT;
	END_VAR

	VAR_OUTPUT
		SIZE2 :	INT;
	END_VAR

	VAR
		a :	INT;
		b :	WORD;
		i :	INT;
		i2 :	INT;
		i3 :	INT;
		c :	INT;
		BASE64 :	STRING := 'ABCDEFGHIJKLMNOPQRSTUVWXYZabcdefghijklmnopqrstuvwxyz0123456789+/';
	END_VAR

	IF SIZE1 <= 0 THEN
		SIZE2 := 0;
		RETURN;
	END_IF;
	c := SIZE1 - 1;
	i2 := 0;
	a := 0;
	b := WORD#0;
	FOR i := 0 TO c DO
		b := SHL(b,8) OR BYTE_TO_WORD(BUF1[i]);
		a := a + 8;
		WHILE a >= 6 DO
			a := a - 6;
			buf2[i2] := INT_TO_BYTE(GET_CHAR(BASE64,WORD_TO_INT(SHR(b,a)) + 1));
			i2 := i2 + 1;
			b := b AND NOT SHL(WORD#16#FFFF,a);
		END_WHILE;
	END_FOR;
	IF a > 0 THEN
		buf2[i2] := INT_TO_BYTE(GET_CHAR(BASE64,WORD_TO_INT(SHL(b,6 - a)) + 1));
		i2 := i2 + 1;
		i3 := i2 + WORD_TO_INT(NOT INT_TO_WORD(i2) AND WORD#2#11);
		FOR i := i2 TO i3 DO
			buf2[i] := BYTE#61;
		END_FOR;
		SIZE2 := i3 + 1;
	ELSE
		SIZE2 := i2;
	END_IF;

END_FUNCTION_BLOCK

PROGRAM program0
  VAR
	BUF1  :	oscat_aB0_63;
	BUF2  :	oscat_aB0_47;

	SIZE1 :	INT;

	SIZE2 :	INT;
	func_block : BASE64_ENCODE_STREAM;
  END_VAR
	func_block.BUF1 :=BUF1 ;
	func_block.BUF2 :=BUF2 ;
	func_block.SIZE1:=SIZE1;
	func_block();
	BUF1 := func_block.BUF1;
	BUF2 := func_block.BUF2;
	SIZE2 := func_block.SIZE2;
END_PROGRAM

CONFIGURATION Config0
  RESOURCE Res0 ON PLC
    TASK task0(INTERVAL := T#20ms,PRIORITY := 0);
    PROGRAM instance0 WITH task0 : program0;
  END_RESOURCE
END_CONFIGURATION

(* ---- BIN_TO_BYTE.ST ---- *)
TYPE
  oscat_STRING12              : STRING(12);
END_TYPE

FUNCTION_BLOCK BIN_TO_BYTE_Block
	VAR_INPUT
		BIN :	oscat_STRING12;
	END_VAR

	VAR_OUTPUT
		BIN_TO_BYTE :	BYTE;
	END_VAR

	VAR
		i :	INT;
		stop :	INT;
		X :	INT;
	END_VAR

	BIN_TO_BYTE := BYTE#0;
	stop := LEN(bin);
	FOR I := 1 TO LEN(BIN) DO
		X := GET_CHAR(BIN,I);
		(* calculate the value of the digit *)
		IF X = 48 THEN
			BIN_TO_BYTE := SHL_BYTE(BIN_TO_BYTE,1);
		ELSIF X = 49 THEN
			BIN_TO_BYTE := SHL_BYTE(BIN_TO_BYTE,1) OR BYTE#1;
		END_IF;
	END_FOR;

END_FUNCTION_BLOCK

PROGRAM program0
  VAR
    LocalVar0 : oscat_STRING12;
	LocalOUT  : BYTE;
	func_block : BIN_TO_BYTE_Block;
  END_VAR
	func_block.BIN := LocalVar0;
	func_block();
	LocalOUT := func_block.BIN_TO_BYTE;

END_PROGRAM

CONFIGURATION Config0
  RESOURCE Res0 ON PLC
    TASK task0(INTERVAL := T#20ms,PRIORITY := 0);
    PROGRAM instance0 WITH task0 : program0;
  END_RESOURCE
END_CONFIGURATION

(* ---- BLIND_ACTUATOR.ST ---- *)
FUNCTION_BLOCK INTERLOCK_Block

	VAR_INPUT
		I1 :	BOOL;
		I2 :	BOOL;
		TL :	TIME;
	END_VAR

	VAR_OUTPUT
		Q1 :	BOOL;
		Q2 :	BOOL;
	END_VAR

	VAR
		T1 :	TOF;
		T2 :	TOF;
	END_VAR

	T1(IN := I1, PT := TL);
	T2(IN := I2, PT := TL);

	Q1 := I1 AND NOT t2.Q;
	Q2 := I2 AND NOT t1.Q;

END_FUNCTION_BLOCK

FUNCTION TIME_TO_UDINT2:UDINT
	VAR_INPUT
		X :	TIME;
	END_VAR

	TIME_TO_UDINT2 := DINT_TO_UDINT(TIME_TO_DINT(X));
END_FUNCTION

FUNCTION_BLOCK T_PLC_MS_block
	VAR_OUTPUT
		T_PLC_MS :	UDINT;
	END_VAR

	VAR_EXTERNAL
		PLC_TICKS_PER_SEC :	INT;
		PLC_SYS_TICK_CNT :	DINT;
	END_VAR

	VAR
		debug :	BOOL;(*Debug-Mode ON / OFF*)
		N :	INT;(*Debug-Faktor*)
		Offset :	UDINT;(*Debug-Offset*)
		temp :	DWORD := DWORD#1;(*Debug-Offset*)
		mode :	BOOL;(*modus*)
		faktor :	UDINT;(*Systemtakt-Faktor*)
		init :	BOOL;
		v_plc_ticks_per_sec :	UDINT;
		base :	UDINT := UDINT#1000;
	END_VAR

	IF init = FALSE THEN
		v_plc_ticks_per_sec := INT_TO_UDINT(PLC_TICKS_PER_SEC);
		IF v_plc_ticks_per_sec = UDINT#1024 THEN
			faktor := UDINT#1;
			mode := FALSE;
		ELSIF v_plc_ticks_per_sec > UDINT#0 THEN
			IF v_plc_ticks_per_sec <= base THEN
				faktor := base / v_plc_ticks_per_sec;
				mode := FALSE;
			ELSE
				faktor := v_plc_ticks_per_sec / base;
				mode := TRUE;
			END_IF;
		ELSE
			faktor := UDINT#1;
		END_IF;
		init := TRUE;
	END_IF;

	IF mode THEN
		T_PLC_MS := DINT_TO_UDINT(PLC_SYS_TICK_CNT) / faktor;
	ELSE
		T_PLC_MS := DINT_TO_UDINT(PLC_SYS_TICK_CNT) * faktor;
	END_IF;

	IF debug THEN
		T_PLC_MS := (DWORD_TO_UDINT(SHL(UDINT_TO_DWORD(T_PLC_MS),N) OR SHL(temp,N)) - UDINT#1) + Offset;
	END_IF;
END_FUNCTION_BLOCK

FUNCTION FRMP_B:BYTE
	VAR_INPUT
		START :	BYTE;
		DIR :	BOOL;
		TD :	TIME;
		TR :	TIME;
	END_VAR

	IF TD < TR THEN
		FRMP_B := MIN(UDINT_TO_BYTE(DWORD_TO_UDINT(SHL(TIME_TO_DWORD(TD), 8)) / TIME_TO_UDINT2(TR)), SEL(DIR, START, USINT_TO_BYTE(USINT#255 - BYTE_TO_USINT(START))));
		IF DIR THEN
			FRMP_B := USINT_TO_BYTE(BYTE_TO_USINT(START) + BYTE_TO_USINT(FRMP_B));
		ELSE
			FRMP_B := USINT_TO_BYTE(BYTE_TO_USINT(START) - BYTE_TO_USINT(FRMP_B));
		END_IF;
	ELSE
		FRMP_B := SEL(DIR, BYTE#0, BYTE#255);
	END_IF;
END_FUNCTION

FUNCTION_BLOCK _RMP_B
	VAR_INPUT
		DIR :	BOOL;
		E :	BOOL := TRUE;
		TR :	TIME;
	END_VAR

	VAR_IN_OUT
		RMP :	BYTE;
	END_VAR

	VAR
		T_PLC_MS :	T_PLC_MS_block;
		tx :	TIME;
		tl :	TIME;
		tn :	TIME;
		init :	BOOL;
		last_dir :	BOOL;
		start :	BYTE;
	END_VAR

	T_PLC_MS();
	tx := UDINT_TO_TIME(T_PLC_MS.T_PLC_MS);

	IF E AND init AND (dir = last_dir) AND (RMP <> SEL(DIR, BYTE#0, BYTE#255)) AND TR = tn THEN
		RMP := FRMP_B(start, DIR, tx - tl, TR);
	ELSE
		init := TRUE;
		tl := tx;
		tn := tr;
		start := RMP;
	END_IF;
	last_dir := dir;
END_FUNCTION_BLOCK

FUNCTION_BLOCK RMP_B_Block

	VAR_INPUT
		SET :	BOOL;
		PT :	TIME;
		E :	BOOL := TRUE;
		UP :	BOOL := TRUE;
		RST :	BOOL;
	END_VAR

	VAR_OUTPUT
		OUT :	BYTE;
		BUSY :	BOOL;
		HIGH :	BOOL;
		LOW :	BOOL;
	END_VAR

	VAR
		rmp :	_RMP_B;
	END_VAR

	rmp(dir := UP, E := E, TR := PT, RMP := out);
	out := rmp.RMP;

	IF RST THEN
		out := BYTE#0;
	ELSIF SET THEN
		out := BYTE#255;
	END_IF;

low := out = BYTE#0;
high := out = BYTE#255;
busy := NOT (low OR high) AND E;

END_FUNCTION_BLOCK

FUNCTION_BLOCK BLIND_ACTUATOR_Block

	VAR_INPUT
		UP :	BOOL;
		DN :	BOOL;
		S_IN :	BYTE;
		T_UD :	TIME := T#10s;
		T_ANGLE :	TIME := T#3s;
		T_LOCKOUT :	TIME := t#100ms;
	END_VAR

	VAR_OUTPUT
		POS :	BYTE;
		ANG :	BYTE;
		QU :	BOOL;
		QD :	BOOL;
		STATUS :	BYTE;
	END_VAR

	VAR
		position :	RMP_B_Block;
		angle :	RMP_B_Block;
		lock :	INTERLOCK_Block;
	END_VAR

	lock(i1 := UP, I2 := DN, TL := T_lockout);

	angle(e := lock.Q1 OR lock.Q2, UP := lock.Q1, PT := T_Angle);
	position(e := lock.Q1 AND angle.high OR lock.Q2 AND angle.low, up := lock.Q1, PT := T_UD);

	pos := position.Out;
	ang := angle.Out;

	QU := lock.Q1;
	QD := lock.Q2;

	IF UP AND DN THEN
		status := BYTE#1;
	ELSIF UP THEN
		status := BYTE#121;
	ELSIF DN THEN
		status := BYTE#122;
	ELSE
		status := S_IN;
	END_IF;

END_FUNCTION_BLOCK

PROGRAM program0
	VAR
		UP :	BOOL;
		DN :	BOOL;
		S_IN :	BYTE;
		T_UD :	TIME := T#10s;
		T_ANGLE :	TIME := T#3s;
		T_LOCKOUT :	TIME := t#100ms;
		POS :	BYTE;
		ANG :	BYTE;
		QU :	BOOL;
		QD :	BOOL;
		func_block : BLIND_ACTUATOR_Block;
	END_VAR
	func_block.UP := UP;
	func_block.DN := DN;
	func_block.S_IN := S_IN ;
	func_block.T_UD := T_UD;
	func_block.T_ANGLE := T_ANGLE;
	func_block.T_LOCKOUT := T_LOCKOUT;
	func_block();
	POS  := func_block.POS;
	ANG  := func_block.ANG;
	QU  := func_block.QU;
	QD  := func_block.QD;
END_PROGRAM

CONFIGURATION Config0
	VAR_GLOBAL
		PLC_TICKS_PER_SEC :	INT;
		PLC_SYS_TICK_CNT :	DINT;
	END_VAR
  	RESOURCE Res0 ON PLC
    	TASK task0(INTERVAL := T#20ms,PRIORITY := 0);
    	PROGRAM instance0 WITH task0 : program0;
  	END_RESOURCE
END_CONFIGURATION

(* ---- BLIND_CONTROL.ST ---- *)
FUNCTION_BLOCK INTERLOCK_Block

	VAR_INPUT
		I1 :	BOOL;
		I2 :	BOOL;
		TL :	TIME;
	END_VAR

	VAR_OUTPUT
		Q1 :	BOOL;
		Q2 :	BOOL;
	END_VAR

	VAR
		T1 :	TOF;
		T2 :	TOF;
	END_VAR

	T1(IN := I1, PT := TL);
	T2(IN := I2, PT := TL);

	Q1 := I1 AND NOT t2.Q;
	Q2 := I2 AND NOT t1.Q;

END_FUNCTION_BLOCK

FUNCTION TIME_TO_UDINT2:UDINT
	VAR_INPUT
		X :	TIME;
	END_VAR

	TIME_TO_UDINT2 := DINT_TO_UDINT(TIME_TO_DINT(X));
END_FUNCTION

FUNCTION_BLOCK T_PLC_MS_block
	VAR_OUTPUT
		T_PLC_MS :	UDINT;
	END_VAR

	VAR_EXTERNAL
		PLC_TICKS_PER_SEC :	INT;
		PLC_SYS_TICK_CNT :	DINT;
	END_VAR

	VAR
		debug :	BOOL;(*Debug-Mode ON / OFF*)
		N :	INT;(*Debug-Faktor*)
		Offset :	UDINT;(*Debug-Offset*)
		temp :	DWORD := DWORD#1;(*Debug-Offset*)
		mode :	BOOL;(*modus*)
		faktor :	UDINT;(*Systemtakt-Faktor*)
		init :	BOOL;
		v_plc_ticks_per_sec :	UDINT;
		base :	UDINT := UDINT#1000;
	END_VAR

	IF init = FALSE THEN
		v_plc_ticks_per_sec := INT_TO_UDINT(PLC_TICKS_PER_SEC);
		IF v_plc_ticks_per_sec = UDINT#1024 THEN
			faktor := UDINT#1;
			mode := FALSE;
		ELSIF v_plc_ticks_per_sec > UDINT#0 THEN
			IF v_plc_ticks_per_sec <= base THEN
				faktor := base / v_plc_ticks_per_sec;
				mode := FALSE;
			ELSE
				faktor := v_plc_ticks_per_sec / base;
				mode := TRUE;
			END_IF;
		ELSE
			faktor := UDINT#1;
		END_IF;
		init := TRUE;
	END_IF;

	IF mode THEN
		T_PLC_MS := DINT_TO_UDINT(PLC_SYS_TICK_CNT) / faktor;
	ELSE
		T_PLC_MS := DINT_TO_UDINT(PLC_SYS_TICK_CNT) * faktor;
	END_IF;

	IF debug THEN
		T_PLC_MS := (DWORD_TO_UDINT(SHL(UDINT_TO_DWORD(T_PLC_MS),N) OR SHL(temp,N)) - UDINT#1) + Offset;
	END_IF;
END_FUNCTION_BLOCK

FUNCTION FRMP_B:BYTE
	VAR_INPUT
		START :	BYTE;
		DIR :	BOOL;
		TD :	TIME;
		TR :	TIME;
	END_VAR

	IF TD < TR THEN
		FRMP_B := MIN(UDINT_TO_BYTE(DWORD_TO_UDINT(SHL(TIME_TO_DWORD(TD), 8)) / TIME_TO_UDINT2(TR)), SEL(DIR, START, USINT_TO_BYTE(USINT#255 - BYTE_TO_USINT(START))));
		IF DIR THEN
			FRMP_B := USINT_TO_BYTE(BYTE_TO_USINT(START) + BYTE_TO_USINT(FRMP_B));
		ELSE
			FRMP_B := USINT_TO_BYTE(BYTE_TO_USINT(START) - BYTE_TO_USINT(FRMP_B));
		END_IF;
	ELSE
		FRMP_B := SEL(DIR, BYTE#0, BYTE#255);
	END_IF;
END_FUNCTION

FUNCTION_BLOCK _RMP_B
	VAR_INPUT
		DIR :	BOOL;
		E :	BOOL := TRUE;
		TR :	TIME;
	END_VAR

	VAR_IN_OUT
		RMP :	BYTE;
	END_VAR

	VAR
		T_PLC_MS :	T_PLC_MS_block;
		tx :	TIME;
		tl :	TIME;
		tn :	TIME;
		init :	BOOL;
		last_dir :	BOOL;
		start :	BYTE;
	END_VAR

	T_PLC_MS();
	tx := UDINT_TO_TIME(T_PLC_MS.T_PLC_MS);

	IF E AND init AND (dir = last_dir) AND (RMP <> SEL(DIR, BYTE#0, BYTE#255)) AND TR = tn THEN
		RMP := FRMP_B(start, DIR, tx - tl, TR);
	ELSE
		init := TRUE;
		tl := tx;
		tn := tr;
		start := RMP;
	END_IF;
	last_dir := dir;
END_FUNCTION_BLOCK

FUNCTION_BLOCK RMP_B_Block

	VAR_INPUT
		SET :	BOOL;
		PT :	TIME;
		E :	BOOL := TRUE;
		UP :	BOOL := TRUE;
		RST :	BOOL;
	END_VAR

	VAR_OUTPUT
		OUT :	BYTE;
		BUSY :	BOOL;
		HIGH :	BOOL;
		LOW :	BOOL;
	END_VAR

	VAR
		rmp :	_RMP_B;
	END_VAR

	rmp(dir := UP, E := E, TR := PT, RMP := out);
	out := rmp.RMP;

	IF RST THEN
		out := BYTE#0;
	ELSIF SET THEN
		out := BYTE#255;
	END_IF;

low := out = BYTE#0;
high := out = BYTE#255;
busy := NOT (low OR high) AND E;

END_FUNCTION_BLOCK

FUNCTION_BLOCK BLIND_ACTUATOR_Block

	VAR_INPUT
		UP :	BOOL;
		DN :	BOOL;
		S_IN :	BYTE;
		T_UD :	TIME := T#10s;
		T_ANGLE :	TIME := T#3s;
		T_LOCKOUT :	TIME := t#100ms;
	END_VAR

	VAR_OUTPUT
		POS :	BYTE;
		ANG :	BYTE;
		QU :	BOOL;
		QD :	BOOL;
		STATUS :	BYTE;
	END_VAR

	VAR
		position :	RMP_B_Block;
		angle :	RMP_B_Block;
		lock :	INTERLOCK_Block;
	END_VAR

	lock(i1 := UP, I2 := DN, TL := T_lockout);

	angle(e := lock.Q1 OR lock.Q2, UP := lock.Q1, PT := T_Angle);
	position(e := lock.Q1 AND angle.high OR lock.Q2 AND angle.low, up := lock.Q1, PT := T_UD);

	pos := position.Out;
	ang := angle.Out;

	QU := lock.Q1;
	QD := lock.Q2;

	IF UP AND DN THEN
		status := BYTE#1;
	ELSIF UP THEN
		status := BYTE#121;
	ELSIF DN THEN
		status := BYTE#122;
	ELSE
		status := S_IN;
	END_IF;

END_FUNCTION_BLOCK

FUNCTION _BYTE_TO_INT:INT
	VAR_INPUT
		IN :	BYTE;
	END_VAR

	_BYTE_TO_INT := USINT_TO_INT(BYTE_TO_USINT(IN));
END_FUNCTION

FUNCTION_BLOCK BLIND_CONTROL_Block

	VAR_INPUT
		UP :	BOOL;
		DN :	BOOL;
		S_IN :	BYTE;
		PI :	BYTE;
		AI :	BYTE;
		T_UD :	TIME;
		T_ANGLE :	TIME;
		SENS :	BYTE := 5;
		T_LOCKOUT :	TIME := T#100ms;
	END_VAR

	VAR_OUTPUT
		POS :	BYTE;
		ANG :	BYTE;
		MU :	BOOL;
		MD :	BOOL;
		STATUS :	BYTE;
	END_VAR

	VAR
		act :	BLIND_ACTUATOR_Block;
		delta :	BYTE;
		bTimeTest :	BOOL;
		iPos :	BYTE;
		iAngel :	BYTE;
	END_VAR

	IF bTimeTest THEN
		PI:=iPos;
		AI:=iAngel;
		UP:=TRUE;
		DN:=TRUE;
	END_IF;

	act(T_UD:=T_UD, T_ANGLE:=T_ANGLE, T_lockout := T_Lockout);

	IF UP AND DN THEN
		IF _BYTE_TO_INT(act.pos) < _BYTE_TO_INT(pi) - _BYTE_TO_INT(delta) THEN
			act.UP := TRUE;
			act.DN := FALSE;
			delta := BYTE#0;
			STATUS := BYTE#121;
		ELSIF _BYTE_TO_INT(act.pos) > _BYTE_TO_INT(pi) + _BYTE_TO_INT(delta) THEN
			act.UP := FALSE;
			act.DN := TRUE;
			delta := BYTE#0;
			STATUS := BYTE#122;
		ELSIF _BYTE_TO_INT(act.ang) < _BYTE_TO_INT(ai) - _BYTE_TO_INT(delta) AND T_angle > T#100ms THEN
			act.UP := TRUE;
			act.DN := FALSE;
			delta := SHR(sens,2);
			STATUS := BYTE#123;
		ELSIF _BYTE_TO_INT(act.ang) > _BYTE_TO_INT(ai) + _BYTE_TO_INT(delta) AND T_angle > T#100ms THEN
			act.UP := FALSE;
			act.DN := TRUE;
			delta := SHR(sens,2);
			STATUS := BYTE#124;
		ELSE
			act.UP := FALSE;
			act.DN := FALSE;
			delta := sens;
			STATUS := S_IN;
		END_IF;
	ELSE
		act.UP := UP;
		act.DN := DN;
		STATUS := S_IN;
	END_IF;

	act(T_UD:=T_UD, T_ANGLE:=T_ANGLE, T_lockout := T_Lockout);
	pos := act.pos;
	ang := act.ang;
	MU := act.QU;
	md := act.QD;
	status := act.status;

END_FUNCTION_BLOCK

PROGRAM program0
	VAR
		UP :	BOOL;
		DN :	BOOL;
		S_IN :	BYTE;
		PI :	BYTE;
		AI :	BYTE;
		T_UD :	TIME;
		T_ANGLE :	TIME;
		SENS :	BYTE := 5;
		T_LOCKOUT :	TIME := T#100ms;
		POS :	BYTE;
		ANG :	BYTE;
		MU :	BOOL;
		MD :	BOOL;
		STATUS :	BYTE;
		func_block : BLIND_CONTROL_Block;
	END_VAR
	func_block.UP := UP;
	func_block.DN := DN;
	func_block.S_IN := S_IN ;
	func_block.PI    := PI    ;
	func_block.AI := AI;
	func_block.T_UD := T_UD ;
	func_block.T_ANGLE    := T_ANGLE    ;
	func_block.SENS := SENS;
	func_block.T_LOCKOUT := T_LOCKOUT;
	func_block();
	POS  := func_block.POS;
	ANG  := func_block.ANG;
	MU  := func_block.MU;
	MD  := func_block.MD;
	STATUS  := func_block.STATUS;
END_PROGRAM

CONFIGURATION Config0
	VAR_GLOBAL
		PLC_TICKS_PER_SEC :	INT;
		PLC_SYS_TICK_CNT :	DINT;
	END_VAR
  	RESOURCE Res0 ON PLC
    	TASK task0(INTERVAL := T#20ms,PRIORITY := 0);
    	PROGRAM instance0 WITH task0 : program0;
  	END_RESOURCE
END_CONFIGURATION

(* ---- BLIND_CONTROL_S.ST ---- *)
FUNCTION UDINT_TO_TIME2:TIME

	VAR_INPUT
		IN :	UDINT;
	END_VAR

	UDINT_TO_TIME2 := DINT_TO_TIME(UDINT_TO_DINT(IN));

END_FUNCTION

FUNCTION_BLOCK T_PLC_MS_block
	VAR_OUTPUT
		T_PLC_MS :	UDINT;
	END_VAR

	VAR_EXTERNAL
		PLC_TICKS_PER_SEC :	INT;
		PLC_SYS_TICK_CNT :	DINT;
	END_VAR

	VAR
		debug :	BOOL;(*Debug-Mode ON / OFF*)
		N :	INT;(*Debug-Faktor*)
		Offset :	UDINT;(*Debug-Offset*)
		temp :	DWORD := DWORD#1;(*Debug-Offset*)
		mode :	BOOL;(*modus*)
		faktor :	UDINT;(*Systemtakt-Faktor*)
		init :	BOOL;
		v_plc_ticks_per_sec :	UDINT;
		base :	UDINT := UDINT#1000;
	END_VAR

	IF init = FALSE THEN
		v_plc_ticks_per_sec := INT_TO_UDINT(PLC_TICKS_PER_SEC);
		IF v_plc_ticks_per_sec = UDINT#1024 THEN
			faktor := UDINT#1;
			mode := FALSE;
		ELSIF v_plc_ticks_per_sec > UDINT#0 THEN
			IF v_plc_ticks_per_sec <= base THEN
				faktor := base / v_plc_ticks_per_sec;
				mode := FALSE;
			ELSE
				faktor := v_plc_ticks_per_sec / base;
				mode := TRUE;
			END_IF;
		ELSE
			faktor := UDINT#1;
		END_IF;
		init := TRUE;
	END_IF;

	IF mode THEN
		T_PLC_MS := DINT_TO_UDINT(PLC_SYS_TICK_CNT) / faktor;
	ELSE
		T_PLC_MS := DINT_TO_UDINT(PLC_SYS_TICK_CNT) * faktor;
	END_IF;

	IF debug THEN
		T_PLC_MS := (DWORD_TO_UDINT(SHL(UDINT_TO_DWORD(T_PLC_MS),N) OR SHL(temp,N)) - UDINT#1) + Offset;
	END_IF;
END_FUNCTION_BLOCK

FUNCTION TIME_TO_UDINT2:UDINT
	VAR_INPUT
		X :	TIME;
	END_VAR

	TIME_TO_UDINT2 := DINT_TO_UDINT(TIME_TO_DINT(X));
END_FUNCTION

FUNCTION FRMP_B:BYTE
	VAR_INPUT
		START :	BYTE;
		DIR :	BOOL;
		TD :	TIME;
		TR :	TIME;
	END_VAR

	IF TD < TR THEN
		FRMP_B := MIN(UDINT_TO_BYTE(DWORD_TO_UDINT(SHL(TIME_TO_DWORD(TD), 8)) / TIME_TO_UDINT2(TR)), SEL(DIR, START, USINT_TO_BYTE(USINT#255 - BYTE_TO_USINT(START))));
		IF DIR THEN
			FRMP_B := USINT_TO_BYTE(BYTE_TO_USINT(START) + BYTE_TO_USINT(FRMP_B));
		ELSE
			FRMP_B := USINT_TO_BYTE(BYTE_TO_USINT(START) - BYTE_TO_USINT(FRMP_B));
		END_IF;
	ELSE
		FRMP_B := SEL(DIR, BYTE#0, BYTE#255);
	END_IF;
END_FUNCTION

FUNCTION_BLOCK _RMP_B
	VAR_INPUT
		DIR :	BOOL;
		E :	BOOL := TRUE;
		TR :	TIME;
	END_VAR

	VAR_IN_OUT
		RMP :	BYTE;
	END_VAR

	VAR
		T_PLC_MS :	T_PLC_MS_block;
		tx :	TIME;
		tl :	TIME;
		tn :	TIME;
		init :	BOOL;
		last_dir :	BOOL;
		start :	BYTE;
	END_VAR

	T_PLC_MS();
	tx := UDINT_TO_TIME(T_PLC_MS.T_PLC_MS);

	IF E AND init AND (dir = last_dir) AND (RMP <> SEL(DIR, BYTE#0, BYTE#255)) AND TR = tn THEN
		RMP := FRMP_B(start, DIR, tx - tl, TR);
	ELSE
		init := TRUE;
		tl := tx;
		tn := tr;
		start := RMP;
	END_IF;
	last_dir := dir;
END_FUNCTION_BLOCK

FUNCTION_BLOCK TREND_DW
	VAR_INPUT
		X :	DWORD;
	END_VAR
	VAR_OUTPUT
		Q :	BOOL;
		TU :	BOOL;
		TD :	BOOL;
		D :	DWORD;
	END_VAR

	VAR
		LAST_X :	DWORD;
	END_VAR

	IF X > last_X THEN
		TU := TRUE;
		TD := FALSE;
		D := UDINT_TO_DWORD(DWORD_TO_UDINT(X) - DWORD_TO_UDINT(last_X));
		Q := TRUE;
	ELSIF X < last_X THEN
		TD := TRUE;
		TU := FALSE;
		D := UDINT_TO_DWORD(DWORD_TO_UDINT(last_X) - DWORD_TO_UDINT(X));
		Q := FALSE;
	ELSE
		TU := FALSE;
		TD := FALSE;
		D := DWORD#0;
	END_IF;
	last_X := X;
END_FUNCTION_BLOCK

FUNCTION_BLOCK _RMP_NEXT
	VAR_INPUT
		E :	BOOL := TRUE;
		IN :	BYTE;
		TR :	TIME;
		TF :	TIME;
		TL :	TIME;
	END_VAR

	VAR_OUTPUT
		DIR :	BOOL;
		UP :	BOOL;
		DN :	BOOL;
	END_VAR

	VAR_IN_OUT
		OUT :	BYTE;
	END_VAR
	VAR
		rmx :	_RMP_B;
		dirx :	TREND_DW;
		t_lock :	TP;
		xen :	BOOL;
		xdir :	BOOL;
	END_VAR

	dirx(X := BYTE_TO_DWORD(in));

	t_lock(in := FALSE, pt := TL);

	IF dirx.TU AND (OUT < IN) THEN
		IF NOT xdir AND xen THEN t_lock(in := TRUE); END_IF;
		xen := TRUE;
		xdir := TRUE;
	ELSIF dirx.TD AND (OUT > IN) THEN
		IF xdir AND xen THEN t_lock(in := TRUE); END_IF;
		xen := TRUE;
		xdir := FALSE;
	ELSIF xen THEN
		IF (xdir AND (out >= in)) OR (NOT xdir AND (out <= in)) THEN
			xen := FALSE;
			IF tl > t#0s THEN t_lock(IN := TRUE); END_IF;
		END_IF;
	END_IF;

	IF NOT t_lock.Q AND xen THEN
		UP := XDIR;
		DIR := XDIR;
		DN := NOT XDIR;
	ELSE
		UP := FALSE;
		DN := FALSE;
	END_IF;

	rmx(rmp := OUT, E := E AND (UP OR DN) , dir := DIR, tr := SEL(dir, TF, TR));
	OUT := rmx.RMP;
END_FUNCTION_BLOCK

FUNCTION _BYTE_TO_INT:INT
	VAR_INPUT
		IN :	BYTE;
	END_VAR

	_BYTE_TO_INT := USINT_TO_INT(BYTE_TO_USINT(IN));
END_FUNCTION

FUNCTION_BLOCK BLIND_CONTROL_S_Block

	VAR_INPUT
		UP :	BOOL;
		DN :	BOOL;
		S_IN :	BYTE := BYTE#125;
		PI :	BYTE;
		T_UP :	TIME;
		T_DN :	TIME;
		RU :	BOOL;
		RD :	BOOL;
		T_LOCKOUT :	TIME := T#100ms;
		T_EXT :	TIME;
		EXT_TRIG :	BYTE := BYTE#5;
		R_POS_TOP :	BYTE := BYTE#255;
		R_POS_BOT :	BYTE;
	END_VAR

	VAR_OUTPUT
		POS :	BYTE;
		MU :	BOOL;
		MD :	BOOL;
		STATUS :	BYTE;
	END_VAR

	VAR
		T_PLC_MS :	T_PLC_MS_Block;
		rmp :	_RMP_NEXT;
		tx :	TIME;
		last :	TIME;
		pi_last :	BYTE;
	END_VAR

	T_PLC_MS();
	tx:= UDINT_TO_TIME(T_PLC_MS.T_PLC_MS);

	IF UP  AND NOT DN THEN
		rmp.IN := BYTE#255;
		STATUS := BYTE#121;
	ELSIF DN AND NOT UP THEN
		rmp.IN := BYTE#0;
		STATUS := BYTE#122;
	ELSIF NOT (UP OR DN) THEN
		rmp.IN := PI;
		STATUS := S_IN;
	END_IF;

	rmp(E := UP OR DN, TR := T_UP, TF := T_DN, TL := T_LOCKOUT, OUT := POS);
	pos := rmp.OUT;

	CASE _BYTE_TO_INT(STATUS) OF
		0:
			last := tx;
			PI_last := PI XOR BYTE#255;
			STATUS := BYTE#128;

		121:
			MU := TRUE;
			MD := FALSE;
			IF POS >= USINT_TO_BYTE(USINT#255 - BYTE_TO_USINT(EXT_TRIG)) THEN
				POS := BYTE#255;
				last := tx;
				STATUS := BYTE#129;
			END_IF;

		122:
			MD := TRUE;
			MU := FALSE;
			IF POS <= EXT_TRIG THEN
				POS := BYTE#0;
				last := tx;
				STATUS := BYTE#129;
			END_IF;

		123:
			MD := rmp.DN;
			MU := rmp.UP;
			IF NOT (rmp.DN OR rmp.UP) THEN
				IF POS <= EXT_TRIG THEN
					MD := TRUE;
					last := tx;
					STATUS := BYTE#129;
				ELSIF POS >= USINT_TO_BYTE(USINT#255 - BYTE_TO_USINT(EXT_TRIG)) THEN
					MU := TRUE;
					last := tx;
					STATUS := BYTE#129;
				ELSE
					STATUS := S_IN;
				END_IF;
			END_IF;

		124:
			MD := rmp.DN;
			MU := rmp.UP;
			IF NOT(rmp.DN OR rmp.UP) THEN
				PI_last := PI;
				STATUS := S_IN;
			END_IF;

		127:
			IF (tx - last) >= T_LOCKOUT THEN
					STATUS := S_IN;
			END_IF;

		128:
			MU := TRUE;
			MD := FALSE;
			rmp.IN := BYTE#255;
			IF (tx - last) >= (T_UP +  T_EXT) THEN
				MU := FALSE;
				last := tx;
				STATUS := BYTE#127;
			END_IF;

		129:
			IF (tx - last) >= T_EXT THEN
				MU := FALSE;
				MD := FALSE;
				last := tx;
				STATUS := BYTE#127;
			END_IF;

	ELSE
		MU := FALSE;
		MD := FALSE;
		IF PI <> PI_last THEN
			PI_last := PI;
			rmp.IN := PI;
			STATUS := BYTE#123;
		ELSIF POS = BYTE#0 AND RU THEN
			rmp.IN := R_POS_BOT;
			STATUS := BYTE#124;
		ELSIF pos = BYTE#255 AND RD THEN
			rmp.IN := R_POS_TOP;
			STATUS := BYTE#124;
		ELSE
			STATUS := S_IN;
		END_IF;
	END_CASE;

END_FUNCTION_BLOCK

PROGRAM program0
	VAR
		UP :	BOOL;
		DN :	BOOL;
		S_IN :	BYTE := BYTE#125;
		PI :	BYTE;
		T_UP :	TIME;
		T_DN :	TIME;
		RU :	BOOL;
		RD :	BOOL;
		T_LOCKOUT :	TIME := T#100ms;
		T_EXT :	TIME;
		EXT_TRIG :	BYTE := BYTE#5;
		R_POS_TOP :	BYTE := BYTE#255;
		R_POS_BOT :	BYTE;
		POS :	BYTE;
		MU :	BOOL;
		MD :	BOOL;
		STATUS :	BYTE;
		func_block : BLIND_CONTROL_S_Block;
	END_VAR
	func_block.UP := UP;
	func_block.DN := DN;
	func_block.S_IN := S_IN ;
	func_block.PI    := PI    ;
	func_block.T_UP := T_UP;
	func_block.T_DN := T_DN ;
	func_block.RU    := RU    ;
	func_block.RD := RD;
	func_block.T_LOCKOUT := T_LOCKOUT;
	func_block.T_EXT := T_EXT ;
	func_block.EXT_TRIG    := EXT_TRIG    ;
	func_block.R_POS_TOP := R_POS_TOP;
	func_block.R_POS_BOT := R_POS_BOT ;
	func_block();
	POS  := func_block.POS;
	MU  := func_block.MU;
	MD  := func_block.MD;
	STATUS  := func_block.STATUS;
END_PROGRAM

CONFIGURATION Config0
	VAR_GLOBAL
		PLC_TICKS_PER_SEC :	INT;
		PLC_SYS_TICK_CNT :	DINT;
	END_VAR
  	RESOURCE Res0 ON PLC
    	TASK task0(INTERVAL := T#20ms,PRIORITY := 0);
    	PROGRAM instance0 WITH task0 : program0;
  	END_RESOURCE
END_CONFIGURATION

(* ---- BLIND_INPUT.ST ---- *)
FUNCTION UDINT_TO_TIME2:TIME

	VAR_INPUT
		IN :	UDINT;
	END_VAR

	UDINT_TO_TIME2 := DINT_TO_TIME(UDINT_TO_DINT(IN));

END_FUNCTION

FUNCTION_BLOCK T_PLC_MS_block
	VAR_OUTPUT
		T_PLC_MS :	UDINT;
	END_VAR

	VAR_EXTERNAL
		PLC_TICKS_PER_SEC :	INT;
		PLC_SYS_TICK_CNT :	DINT;
	END_VAR

	VAR
		debug :	BOOL;(*Debug-Mode ON / OFF*)
		N :	INT;(*Debug-Faktor*)
		Offset :	UDINT;(*Debug-Offset*)
		temp :	DWORD := DWORD#1;(*Debug-Offset*)
		mode :	BOOL;(*modus*)
		faktor :	UDINT;(*Systemtakt-Faktor*)
		init :	BOOL;
		v_plc_ticks_per_sec :	UDINT;
		base :	UDINT := UDINT#1000;
	END_VAR

	IF init = FALSE THEN
		v_plc_ticks_per_sec := INT_TO_UDINT(PLC_TICKS_PER_SEC);
		IF v_plc_ticks_per_sec = UDINT#1024 THEN
			faktor := UDINT#1;
			mode := FALSE;
		ELSIF v_plc_ticks_per_sec > UDINT#0 THEN
			IF v_plc_ticks_per_sec <= base THEN
				faktor := base / v_plc_ticks_per_sec;
				mode := FALSE;
			ELSE
				faktor := v_plc_ticks_per_sec / base;
				mode := TRUE;
			END_IF;
		ELSE
			faktor := UDINT#1;
		END_IF;
		init := TRUE;
	END_IF;

	IF mode THEN
		T_PLC_MS := DINT_TO_UDINT(PLC_SYS_TICK_CNT) / faktor;
	ELSE
		T_PLC_MS := DINT_TO_UDINT(PLC_SYS_TICK_CNT) * faktor;
	END_IF;

	IF debug THEN
		T_PLC_MS := (DWORD_TO_UDINT(SHL(UDINT_TO_DWORD(T_PLC_MS),N) OR SHL(temp,N)) - UDINT#1) + Offset;
	END_IF;

END_FUNCTION_BLOCK

FUNCTION_BLOCK CLICK_MODE_Block

	VAR_INPUT
		IN :	BOOL;
		T_LONG :	TIME := T#500ms;
	END_VAR

	VAR_OUTPUT
		SINGLE :	BOOL;
		DOUBLE :	BOOL;
		LONG :	BOOL;
		TP_LONG :	BOOL;
	END_VAR

	VAR
		Timer :	TP;
		cnt :	INT;
		last :	BOOL;
	END_VAR

	timer(in := IN, PT := T_LONG);
	single := FALSE;
	double := FALSE;

	IF timer.Q THEN
		IF NOT in AND last THEN	cnt := cnt + 1; END_IF;
	ELSE
		CASE cnt OF
			1 : single := TRUE;
			2 : double := TRUE;
		END_CASE;
		cnt := 0;
	END_IF;
	last := in;
	TP_LONG := NOT timer.Q AND (NOT LONG) AND IN;
	LONG := NOT timer.Q AND in;

END_FUNCTION_BLOCK

FUNCTION _BYTE_TO_INT:INT
	VAR_INPUT
		IN :	BYTE;
	END_VAR

	_BYTE_TO_INT := USINT_TO_INT(BYTE_TO_USINT(IN));
END_FUNCTION

FUNCTION_BLOCK BLIND_INPUT_Block

	VAR_INPUT
		POS :	BYTE;
		ANG :	BYTE;
		S1 :	BOOL;
		S2 :	BOOL;
		IN :	BOOL;
		PI :	BYTE;
		AI :	BYTE;
		SINGLE_SWITCH :	BOOL;
		CLICK_EN :	BOOL := TRUE;
		CLICK_TIME :	TIME := T#500ms;
		MAX_RUNTIME :	TIME := T#60s;
		MANUAL_TIMEOUT :	TIME := T#1h;
		DEBOUNCE_TIME :	TIME := T#20ms;
		DBL_CLK1 :	BOOL := FALSE;
		DBL_POS1 :	BYTE;
		DBL_ANG1 :	BYTE;
		DBL_CLK2 :	BOOL := FALSE;
		DBL_POS2 :	BYTE := BYTE#255;
		DBL_ANG2 :	BYTE := BYTE#255;
		D1_TOGGLE :	BOOL := TRUE;
		D2_TOGGLE :	BOOL := TRUE;
		MASTER_MODE :	BOOL;
	END_VAR

	VAR_OUTPUT
		QU :	BOOL := TRUE;
		QD :	BOOL := TRUE;
		STATUS :	BYTE;
		PO :	BYTE := BYTE#255;
		AO :	BYTE := BYTE#255;
		D1 :	BOOL;
		D2 :	BOOL;
	END_VAR

	VAR
		s1e :	TOF;
		s2e :	TOF;
		s1d :	CLICK_MODE_Block;
		s2d :	CLICK_MODE_Block;
		dir :	BOOL;
		tx :	TIME;
		last :	TIME;
		T_PLC_MS :	T_PLC_MS_Block;
	END_VAR

	T_PLC_MS();
	tx:= UDINT_TO_TIME(T_PLC_MS.T_PLC_MS);

	s1e(in := S1, pt := DEBOUNCE_TIME);
	s2e(in := S2, pt := DEBOUNCE_TIME);
	s1d(in := (s1e.Q AND NOT SINGLE_SWITCH) OR (s1e.Q AND SINGLE_SWITCH AND dir), t_long := CLICK_TIME);
	s2d(in := (s2e.Q AND NOT SINGLE_SWITCH) OR (s1e.Q AND SINGLE_SWITCH AND NOT dir), t_long := CLICK_TIME);

	IF NOT d1_toggle THEN d1 := FALSE; END_IF;
	IF NOT d2_toggle THEN d2 := FALSE; END_IF;

	IF (s1d.LONG AND s2d.LONG) OR (status = BYTE#139) THEN
	status := BYTE#139;
	IF NOT (s1d.LONG OR s2d.LONG)  THEN status := BYTE#130; END_IF;
	ELSIF s1d.tp_LONG THEN
		status := BYTE#132;
	ELSIF s2d.tp_LONG THEN
		status := BYTE#133;
	ELSIF  s1d.SINGLE THEN
		IF click_en THEN
			IF QU XOR QD THEN
				status := BYTE#131;
			ELSE
				status := BYTE#134;
				last := tx;
				dir := NOT dir;
			END_IF;
		END_IF;
	ELSIF  s2d.SINGLE THEN
		IF click_en THEN
			IF QU XOR QD THEN
				status := BYTE#131;
			ELSE
				status := BYTE#135;
				last := tx;
				dir := NOT dir;
			END_IF;
		END_IF;
	ELSIF in THEN
		status := BYTE#136;
		last := tx;
	ELSIF s1d.DOUBLE THEN
		IF dbl_clk1 THEN
			status := BYTE#137;
			last := tx;
		ELSE
			D1 := NOT D1;
		END_IF;
	ELSIF s2d.DOUBLE THEN
		IF dbl_clk2 THEN
			status := BYTE#138;
			last := tx;
		ELSE
			IF single_switch THEN D1 := NOT D1; ELSE D2 := NOT D2; END_IF;
		END_IF;
	END_IF;

	CASE _BYTE_TO_INT(status) OF
		0:
				status := BYTE#130;

		130:
				IF NOT master_mode THEN
					PO := POS;
					AO := ANG;
				END_IF;
				QU := TRUE;
				QD := TRUE;

		131:
				QU := FALSE;
				QD := FALSE;
				PO := POS;
				AO := ANG;
				IF tx - last >= manual_timeout THEN
					status := BYTE#130;
				END_IF;

		132:
				QU := TRUE;
				QD := FALSE;
				PO := POS; AO := ANG;
				last := tx;
				IF NOT s1d.LONG THEN status := BYTE#131; dir := NOT dir; END_IF;

		133:
				QU := FALSE;
				QD := TRUE;
				PO := POS; AO := ANG;
				last := tx;
				IF NOT s2d.LONG THEN	status := BYTE#131; dir := NOT dir; END_IF;

		134:
				QU := TRUE;
				QD := FALSE;
				PO := POS; AO := ANG;
				IF tx - last >= max_runtime THEN status := BYTE#131; END_IF;

		135:
				QU := FALSE;
				QD := TRUE;
				PO := POS; AO := ANG;
				IF tx - last >= max_runtime THEN status := BYTE#131;	END_IF;

		136:
				QU := TRUE;
				QD := TRUE;
				PO := PI; AO := AI;
				IF tx-last >= max_runtime THEN status := BYTE#130; END_IF;

		137:
				QU := TRUE;
				QD := TRUE;
				PO := DBL_POS1;
				AO := DBL_ANG1;
				IF tx - last >= max_runtime THEN status := BYTE#131; END_IF;

		138:
				QU := TRUE;
				QD := TRUE;
				PO := DBL_POS2;
				AO := DBL_ANG2;
				IF tx - last >= max_runtime THEN status := BYTE#131; END_IF;

		139:
				QU := FALSE;
				QD := FALSE;
				PO := POS;
				AO := ANG;

	END_CASE;

END_FUNCTION_BLOCK

PROGRAM program0
	VAR
		POS :	BYTE;
		ANG :	BYTE;
		S1 :	BOOL;
		S2 :	BOOL;
		IN :	BOOL;
		PI :	BYTE;
		AI :	BYTE;
		SINGLE_SWITCH :	BOOL;
		CLICK_EN :	BOOL := TRUE;
		CLICK_TIME :	TIME := T#500ms;
		MAX_RUNTIME :	TIME := T#60s;
		MANUAL_TIMEOUT :	TIME := T#1h;
		DEBOUNCE_TIME :	TIME := T#20ms;
		DBL_CLK1 :	BOOL := FALSE;
		DBL_POS1 :	BYTE;
		DBL_ANG1 :	BYTE;
		DBL_CLK2 :	BOOL := FALSE;
		DBL_POS2 :	BYTE := BYTE#255;
		DBL_ANG2 :	BYTE := BYTE#255;
		D1_TOGGLE :	BOOL := TRUE;
		D2_TOGGLE :	BOOL := TRUE;
		MASTER_MODE :	BOOL;
		QU :	BOOL := TRUE;
		QD :	BOOL := TRUE;
		STATUS :	BYTE;
		PO :	BYTE := BYTE#255;
		AO :	BYTE := BYTE#255;
		D1 :	BOOL;
		D2 :	BOOL;
		func_block : BLIND_INPUT_Block;
	END_VAR
	func_block.POS := POS;
	func_block.ANG := ANG;
	func_block.S1 := S1 ;
	func_block.S2 := S2;
	func_block.IN := IN;
	func_block.PI := PI;
	func_block.AI := AI;
	func_block.SINGLE_SWITCH := SINGLE_SWITCH;
	func_block.CLICK_EN := CLICK_EN ;
	func_block.CLICK_TIME := CLICK_TIME;
	func_block.MAX_RUNTIME := MAX_RUNTIME;
	func_block.MANUAL_TIMEOUT := MANUAL_TIMEOUT;
	func_block.DEBOUNCE_TIME := DEBOUNCE_TIME;
	func_block.DBL_CLK1 := DBL_CLK1;
	func_block.DBL_POS1 := DBL_POS1 ;
	func_block.DBL_ANG1 := DBL_ANG1;
	func_block.DBL_CLK2 := DBL_CLK2;
	func_block.DBL_POS2 := DBL_POS2;
	func_block.DBL_ANG2 := DBL_ANG2;
	func_block.D1_TOGGLE := D1_TOGGLE ;
	func_block.D2_TOGGLE := D2_TOGGLE;
	func_block.MASTER_MODE := MASTER_MODE;
	func_block();
	QU  := func_block.QU;
	QD  := func_block.QD;
	STATUS  := func_block.STATUS;
	PO  := func_block.PO;
	AO  := func_block.AO;
	D1  := func_block.D1;
	D2  := func_block.D2;
END_PROGRAM

CONFIGURATION Config0
	VAR_GLOBAL
		PLC_TICKS_PER_SEC :	INT;
		PLC_SYS_TICK_CNT :	DINT;
	END_VAR
  	RESOURCE Res0 ON PLC
    	TASK task0(INTERVAL := T#20ms,PRIORITY := 0);
    	PROGRAM instance0 WITH task0 : program0;
  	END_RESOURCE
END_CONFIGURATION

(* ---- BLIND_NIGHT.ST ---- *)
FUNCTION TIME_TO_UDINT2:UDINT
	VAR_INPUT
		X :	TIME;
	END_VAR

	TIME_TO_UDINT2 := DINT_TO_UDINT(TIME_TO_DINT(X));
END_FUNCTION

FUNCTION DT_TO_DATE2:UDINT

	VAR_INPUT
		IN :	UDINT;
	END_VAR

	DT_TO_DATE2 := (IN / UDINT#86400) * UDINT#86400;
END_FUNCTION

FUNCTION DT_TO_TOD2:UDINT
	VAR_INPUT
		IN :	UDINT;
	END_VAR

	DT_TO_TOD2 := (IN MOD UDINT#86400) * UDINT#1000;
END_FUNCTION

FUNCTION_BLOCK BLIND_NIGHT_Block

	VAR_INPUT
		UP :	BOOL;
		DN :	BOOL;
		S_IN :	BYTE;
		PI :	BYTE;
		AI :	BYTE;
		E_NIGHT :	BOOL := TRUE;
		E_DAY :	BOOL := TRUE;
		DTIN :	UDINT;
		SUNRISE :	UDINT;
		SUNSET :	UDINT;
		SUNRISE_OFFSET :	TIME;
		SUNSET_OFFSET :	TIME;
		NIGHT_POSITION :	BYTE;
		NIGHT_ANGLE :	BYTE;
	END_VAR

	VAR_OUTPUT
		QU :	BOOL;
		QD :	BOOL;
		STATUS :	BYTE;
		PO :	BYTE;
		AO :	BYTE;
	END_VAR

	VAR
		night :	BOOL;
		last_night :	UDINT;
		last_day :	UDINT;
	END_VAR

	IF NOT (up AND dn) AND night THEN
		night := FALSE;
	ELSIF (DT_TO_TOD2(dtin) > sunset + TIME_TO_UDINT2(sunset_offset)) AND (last_night < DT_TO_DATE2(dtin)) AND NOT night AND e_night THEN
		night := TRUE;
		last_night := DT_TO_DATE2(dtin);
	ELSIF (DT_TO_TOD2(dtin) > sunrise + TIME_TO_UDINT2(sunrise_offset)) AND (last_day < DT_TO_DATE2(dtin)) AND night AND e_day AND (last_night < DT_TO_DATE2(dtin)) THEN
		night := FALSE;
		last_day := DT_TO_DATE2(dtin);
	END_IF;

	IF UP AND DN AND night THEN
		status := BYTE#141;
		po := night_position;
		ao := night_angle;
	ELSE
		QU := UP;
		QD := DN;
		po := pi;
		ao := ai;
		status := s_in;
	END_IF;

END_FUNCTION_BLOCK

PROGRAM program0
	VAR
		UP :	BOOL;
		DN :	BOOL;
		S_IN :	BYTE;
		PI :	BYTE;
		AI :	BYTE;
		E_NIGHT :	BOOL := TRUE;
		E_DAY :	BOOL := TRUE;
		DTIN :	UDINT;
		SUNRISE :	UDINT;
		SUNSET :	UDINT;
		SUNRISE_OFFSET :	TIME;
		SUNSET_OFFSET :	TIME;
		NIGHT_POSITION :	BYTE;
		NIGHT_ANGLE :	BYTE;
		QU :	BOOL;
		QD :	BOOL;
		STATUS :	BYTE;
		PO :	BYTE;
		AO :	BYTE;

		func_block : BLIND_NIGHT_Block;
	END_VAR
	func_block.UP := UP;
	func_block.DN := DN;
	func_block.S_IN := S_IN ;
	func_block.PI    := PI    ;
	func_block.AI := AI;
	func_block.E_NIGHT := E_NIGHT;
	func_block.E_DAY := E_DAY ;
	func_block.DTIN    := DTIN    ;
	func_block.SUNRISE := SUNRISE;
	func_block.SUNSET := SUNSET;
	func_block.SUNRISE_OFFSET := SUNRISE_OFFSET ;
	func_block.SUNSET_OFFSET    := SUNSET_OFFSET    ;
	func_block.NIGHT_POSITION := NIGHT_POSITION ;
	func_block.NIGHT_ANGLE    := NIGHT_ANGLE    ;

	func_block();
	QU  := func_block.QU;
	QD  := func_block.QD;
	STATUS  := func_block.STATUS;
	PO  := func_block.PO;
	AO  := func_block.AO;
END_PROGRAM

CONFIGURATION Config0
	RESOURCE Res0 ON PLC
		TASK task0(INTERVAL := T#20ms,PRIORITY := 0);
		PROGRAM instance0 WITH task0 : program0;
	END_RESOURCE
END_CONFIGURATION

(* ---- BLIND_SCENE.ST ---- *)
TYPE
	oscat_bsa_X                 : ARRAY [0..2]    OF BYTE;
  	oscat_blind_scene_array     : ARRAY [0..15]   OF oscat_bsa_X := [0, 0, 0, 0, 0, 0, 0, 0, 0, 0, 0, 0, 0, 0, 0, 0];
END_TYPE

FUNCTION _BYTE_TO_INT:INT
	VAR_INPUT
		IN :	BYTE;
	END_VAR

	_BYTE_TO_INT := USINT_TO_INT(BYTE_TO_USINT(IN));
END_FUNCTION

FUNCTION_BLOCK BLIND_SCENE_Block

	VAR_INPUT
		UP :	BOOL;
		DN :	BOOL;
		S_IN :	BYTE;
		PI :	BYTE;
		AI :	BYTE;
		ENABLE :	BOOL;
		SWRITE :	BOOL;
		SCENE :	BYTE;
	END_VAR

	VAR_OUTPUT
		QU :	BOOL;
		QD :	BOOL;
		STATUS :	BYTE;
		PO :	BYTE;
		AO :	BYTE;
	END_VAR

	VAR
		x :	INT;
	END_VAR

	VAR RETAIN
		sx :	oscat_blind_scene_array;
	END_VAR

	x := _BYTE_TO_INT(scene AND BYTE#2#0000_1111);

	IF enable AND (sx[x][2] > BYTE#0) AND UP AND DN THEN
		po := sx[x][0];
		ao := sx[x][1];
		status := INT_TO_BYTE(160 + x);
		QU := TRUE;
		QD := TRUE;
	ELSE
		QU := UP;
		QD := DN;
		status := S_IN;
		po := pi;
		ao := ai;
	END_IF;

	IF swrite THEN
		status := BYTE#176;
		sx[x][0] := pi;
		sx[x][1] := ai;
		IF enable THEN sx[x][2] := BYTE#1; ELSE sx[x][2] := BYTE#0; END_IF;
	END_IF;

END_FUNCTION_BLOCK

PROGRAM program0
	VAR
		UP :	BOOL;
		DN :	BOOL;
		S_IN :	BYTE;
		PI :	BYTE;
		AI :	BYTE;
		ENABLE :	BOOL;
		SWRITE :	BOOL;
		SCENE :	BYTE;
		QU :	BOOL;
		QD :	BOOL;
		STATUS :	BYTE;
		PO :	BYTE;
		AO :	BYTE;

		func_block : BLIND_SCENE_Block;
	END_VAR
	func_block.UP := UP;
	func_block.DN := DN;
	func_block.S_IN := S_IN ;
	func_block.PI    := PI    ;
	func_block.AI := AI;
	func_block.ENABLE := ENABLE;
	func_block.SWRITE := SWRITE ;
	func_block.SCENE := SCENE ;

	func_block();
	QU  := func_block.QU;
	QD  := func_block.QD;
	STATUS  := func_block.STATUS;
	PO  := func_block.PO;
	AO  := func_block.AO;
END_PROGRAM

CONFIGURATION Config0
	RESOURCE Res0 ON PLC
		TASK task0(INTERVAL := T#20ms,PRIORITY := 0);
		PROGRAM instance0 WITH task0 : program0;
	END_RESOURCE
END_CONFIGURATION

(* ---- BLIND_SECURITY.ST ---- *)
FUNCTION_BLOCK BLIND_SECURITY_Block

	VAR_INPUT
		UP :	BOOL;
		DN :	BOOL;
		S_IN :	BYTE;
		PI :	BYTE;
		AI :	BYTE;
		FIRE :	BOOL;
		WIND :	BOOL;
		ALARM :	BOOL;
		DOOR :	BOOL;
		RAIN :	BOOL;
		ALARM_UP :	BOOL := TRUE;
		WIND_UP :	BOOL := TRUE;
		RAIN_UP :	BOOL := TRUE;
	END_VAR

	VAR_OUTPUT
		QU :	BOOL;
		QD :	BOOL;
		STATUS :	BYTE;
		PO :	BYTE;
		AO :	BYTE;
	END_VAR

	IF Fire THEN
		QU := TRUE;
		QD := FALSE;
		status := BYTE#111;
	ELSIF Wind THEN
		QU := Wind_up;
		QD := NOT wind_up;
		status := BYTE#112;
	ELSIF alarm THEN
		QU := Alarm_up;
		QD := NOT Alarm_up;
		status := BYTE#113;
	ELSIF Door THEN
		QU := TRUE;
		QD := FALSE;
		status := BYTE#114;
	ELSIF Rain AND NOT (up XOR dn) THEN
		QU := rain_up;
		QD := NOT rain_up;
		status := BYTE#115;
	ELSE
		QU := UP;
		QD := DN;
		status := S_IN;
		po := pi;
		ao := ai;
	END_IF;

END_FUNCTION_BLOCK

PROGRAM program0
	VAR
		UP :	BOOL;
		DN :	BOOL;
		S_IN :	BYTE;
		PI :	BYTE;
		AI :	BYTE;
		FIRE :	BOOL;
		WIND :	BOOL;
		ALARM :	BOOL;
		DOOR :	BOOL;
		RAIN :	BOOL;
		ALARM_UP :	BOOL := TRUE;
		WIND_UP :	BOOL := TRUE;
		RAIN_UP :	BOOL := TRUE;
		QU :	BOOL;
		QD :	BOOL;
		STATUS :	BYTE;
		PO :	BYTE;
		AO :	BYTE;

		func_block : BLIND_SECURITY_Block;
	END_VAR
	func_block.UP := UP;
	func_block.DN := DN;
	func_block.S_IN := S_IN ;
	func_block.PI    := PI    ;
	func_block.AI := AI;
	func_block.FIRE := FIRE;
	func_block.WIND := WIND ;
	func_block.ALARM := ALARM ;
	func_block.DOOR    := DOOR    ;
	func_block.RAIN := RAIN;
	func_block.ALARM_UP := ALARM_UP;
	func_block.WIND_UP := WIND_UP ;
	func_block.RAIN_UP := RAIN_UP ;

	func_block();
	QU  := func_block.QU;
	QD  := func_block.QD;
	STATUS  := func_block.STATUS;
	PO  := func_block.PO;
	AO  := func_block.AO;
END_PROGRAM

CONFIGURATION Config0
	RESOURCE Res0 ON PLC
		TASK task0(INTERVAL := T#20ms,PRIORITY := 0);
		PROGRAM instance0 WITH task0 : program0;
	END_RESOURCE
END_CONFIGURATION

(* ---- BLIND_SET.ST ---- *)
FUNCTION UDINT_TO_TIME2:TIME

	VAR_INPUT
		IN :	UDINT;
	END_VAR

	UDINT_TO_TIME2 := DINT_TO_TIME(UDINT_TO_DINT(IN));

END_FUNCTION

FUNCTION_BLOCK T_PLC_MS_block
	VAR_OUTPUT
		T_PLC_MS :	UDINT;
	END_VAR

	VAR_EXTERNAL
		PLC_TICKS_PER_SEC :	INT;
		PLC_SYS_TICK_CNT :	DINT;
	END_VAR

	VAR
		debug :	BOOL;(*Debug-Mode ON / OFF*)
		N :	INT;(*Debug-Faktor*)
		Offset :	UDINT;(*Debug-Offset*)
		temp :	DWORD := DWORD#1;(*Debug-Offset*)
		mode :	BOOL;(*modus*)
		faktor :	UDINT;(*Systemtakt-Faktor*)
		init :	BOOL;
		v_plc_ticks_per_sec :	UDINT;
		base :	UDINT := UDINT#1000;
	END_VAR

	IF init = FALSE THEN
		v_plc_ticks_per_sec := INT_TO_UDINT(PLC_TICKS_PER_SEC);
		IF v_plc_ticks_per_sec = UDINT#1024 THEN
			faktor := UDINT#1;
			mode := FALSE;
		ELSIF v_plc_ticks_per_sec > UDINT#0 THEN
			IF v_plc_ticks_per_sec <= base THEN
				faktor := base / v_plc_ticks_per_sec;
				mode := FALSE;
			ELSE
				faktor := v_plc_ticks_per_sec / base;
				mode := TRUE;
			END_IF;
		ELSE
			faktor := UDINT#1;
		END_IF;
		init := TRUE;
	END_IF;

	IF mode THEN
		T_PLC_MS := DINT_TO_UDINT(PLC_SYS_TICK_CNT) / faktor;
	ELSE
		T_PLC_MS := DINT_TO_UDINT(PLC_SYS_TICK_CNT) * faktor;
	END_IF;

	IF debug THEN
		T_PLC_MS := (DWORD_TO_UDINT(SHL(UDINT_TO_DWORD(T_PLC_MS),N) OR SHL(temp,N)) - UDINT#1) + Offset;
	END_IF;

END_FUNCTION_BLOCK

FUNCTION_BLOCK BLIND_SET_Block

	VAR_INPUT
		UP :	BOOL;
		DN :	BOOL;
		S_IN :	INT;
		PI :	BYTE;
		AI :	BYTE;
		IN :	BOOL;
		PX :	BYTE;
		AX :	BYTE;
		OVERRIDE_MANUAL :	BOOL;
		RESTORE_POSITION :	BOOL;
		RESTORE_TIME :	TIME := T#60s;
	END_VAR

	VAR_OUTPUT
		QU :	BOOL;
		QD :	BOOL;
		STATUS :	INT;
		PO :	BYTE;
		AO :	BYTE;
	END_VAR

	VAR
		T_PLC_MS :	T_PLC_MS_Block;
		tx :	TIME;
		ps :	BYTE;
		as :	BYTE;
		last :	TIME;
	END_VAR

	T_PLC_MS();
	tx:= UDINT_TO_TIME(T_PLC_MS.T_PLC_MS);

	IF IN THEN
		IF override_manual OR (UP AND DN) THEN
			status := 178;
		END_IF;
	END_IF;

	CASE STATUS OF
		0:
			status := S_IN;

		178:
			PO := PX;
			AO := AX;
			QU := TRUE;
			QD := TRUE;
			IF NOT in THEN
				STATUS := SEL(RESTORE_POSITION, S_IN, 179);
				last := tx;
			END_IF;

		179:
			PO := ps;
			AO := as;
			IF ((PO = PI) AND (AO = AI))  OR tx - last >= RESTORE_TIME THEN
				status := S_IN;
			END_IF;

	ELSE
		PO := PI;
		ps := PI;
		AO := AI;
		as := AI;
		STATUS := S_IN;
		QU := UP;
		QD := DN;
	END_CASE;

END_FUNCTION_BLOCK

PROGRAM program0
	VAR
		UP :	BOOL;
		DN :	BOOL;
		S_IN :	INT;
		PI :	BYTE;
		AI :	BYTE;
		IN :	BOOL;
		PX :	BYTE;
		AX :	BYTE;
		OVERRIDE_MANUAL :	BOOL;
		RESTORE_POSITION :	BOOL;
		RESTORE_TIME :	TIME := T#60s;
		QU :	BOOL;
		QD :	BOOL;
		STATUS :	INT;
		PO :	BYTE;
		AO :	BYTE;

		func_block : BLIND_SET_Block;
	END_VAR
	func_block.UP := UP;
	func_block.DN := DN;
	func_block.S_IN := S_IN ;
	func_block.PI    := PI    ;
	func_block.AI := AI;
	func_block.IN := IN;
	func_block.PX := PX ;
	func_block.AX := AX ;
	func_block.OVERRIDE_MANUAL    := OVERRIDE_MANUAL    ;
	func_block.RESTORE_POSITION := RESTORE_POSITION;
	func_block.RESTORE_TIME := RESTORE_TIME;

	func_block();
	QU  := func_block.QU;
	QD  := func_block.QD;
	STATUS  := func_block.STATUS;
	PO  := func_block.PO;
	AO  := func_block.AO;
END_PROGRAM

CONFIGURATION Config0
	VAR_GLOBAL
		PLC_TICKS_PER_SEC :	INT;
		PLC_SYS_TICK_CNT :	DINT;
	END_VAR
  	RESOURCE Res0 ON PLC
    	TASK task0(INTERVAL := T#20ms,PRIORITY := 0);
    	PROGRAM instance0 WITH task0 : program0;
  	END_RESOURCE
END_CONFIGURATION

(* ---- BLIND_SHADE.ST ---- *)
TYPE
  oscat_STRING5               : STRING;
  oscat_STRING30              : STRING;
END_TYPE

TYPE oscat_CALENDAR :
	STRUCT
		UTC : UDINT;				(* world time UTC *)
		LDT : UDINT;				(* local time *)
		LDATE : UDINT;				(* local date *)
		LTOD : UDINT;				(* local time of day *)
		YEAR : INT;					(* year of LDATE *)
		MONTH : INT;				(* month of LDATE *)
		DAY : INT;					(* day of LDATE *)
		WEEKDAY : INT;				(* weekday of LDATE *)
		OFFSET : INT;				(* Time Zone Offset for Local time in minutes *)
		DST_EN : BOOL;				(* daylight savings time enable *)
		DST_ON : BOOL;				(* true when daylight savings time os on *)
		NAME : oscat_string5;		(* name of time zone *)
		LANGUAGE : INT;			    (* language number pls see language setup *)
		LONGITUDE : REAL;			(* longitude of current location *)
		LATITUDE : REAL;			(* latitude of current location *)
		SUN_RISE : UDINT;			(* sun_rise for current location *)
		SUN_SET : UDINT;			(* sun_set for current location *)
		SUN_MIDDAY : UDINT;			(* worldtime when sun stands at south position *)
		SUN_HEIGTH : REAL;			(* suns heigth at midday, south position *)
		SUN_HOR : REAL;				(* sun angle horizontal 0 = north in degrees *)
		SUN_VER : REAL;				(* sun angle vertical above horizon in degrees *)
		NIGHT : BOOL;				(* true between sun_set and sun_rise *)
		HOLIDAY : BOOL;				(* true when holiday *)
		HOLY_NAME : oscat_string30;	(* name of holiday *)
		WORK_WEEK : INT;			(* current work week *)
	END_STRUCT;
END_TYPE

FUNCTION DT_TO_TOD2:UDINT
	VAR_INPUT
		IN :	UDINT;
	END_VAR

	DT_TO_TOD2 := (IN MOD UDINT#86400) * UDINT#1000;
END_FUNCTION

FUNCTION TIME_TO_UDINT2:UDINT
	VAR_INPUT
		X :	TIME;
	END_VAR

	TIME_TO_UDINT2 := DINT_TO_UDINT(TIME_TO_DINT(X));
END_FUNCTION

FUNCTION DEG : REAL
	VAR_INPUT
		RAD_IN : REAL;
	END_VAR

	DEG := MODR(57.29577951308232 * RAD_IN, 360.0);
END_FUNCTION

FUNCTION MODR : REAL
	VAR_INPUT
		IN : REAL;
		DIVI : REAL;
	END_VAR

	IF divi = 0.0 THEN
		MODR := 0.0;
	ELSE
		MODR := in - DINT_TO_REAL(FLOOR2(in / divi)) * divi;
	END_IF;
END_FUNCTION

FUNCTION FLOOR2 : DINT
	VAR_INPUT
		x : REAL;
	END_VAR

	FLOOR2 := REAL_TO_DINT(X);
	IF DINT_TO_REAL(FLOOR2) > X THEN
		FLOOR2 := FLOOR2 - DINT#1;
	END_IF;
END_FUNCTION

FUNCTION RAD:REAL

	VAR_INPUT
		DEG1 :	REAL;
	END_VAR

	RAD := MODR(0.0174532925199433 * DEG1 , 6.283185307179586476);

END_FUNCTION

FUNCTION TRUNC_UDINT2:UDINT
	VAR_INPUT
		IN :	REAL;
	END_VAR
	TRUNC_UDINT2 := DINT_TO_UDINT(TRUNC_DINT(IN));
END_FUNCTION

FUNCTION_BLOCK BLIND_SHADE_Block

	VAR_INPUT
		UP :	BOOL;
		DN :	BOOL;
		S_IN :	BYTE;
		PI :	BYTE;
		AI :	BYTE;
		ENABLE :	BOOL;
		SUN :	BOOL;
		SUNRISE_OFFSET :	TIME := T#1h;
		SUNSET_PRESET :	TIME := T#1h;
		DIRECTION :	REAL := 180.0;
		ANGLE_OFFSET :	REAL := 80.0;
		SLAT_WIDTH :	REAL := 80.0;
		SLAT_SPACING :	REAL := 60.0;
		SHADE_DELAY :	TIME := T#60s;
		SHADE_POS :	BYTE;
	END_VAR

	VAR_OUTPUT
		QU :	BOOL;
		QD :	BOOL;
		STATUS :	BYTE;
		PO :	BYTE;
		AO :	BYTE;
	END_VAR

	VAR_IN_OUT
		CX :	oscat_CALENDAR;
	END_VAR

	VAR
		angle :	REAL;
		sun_delay :	TOF;
	END_VAR

	sun_delay(IN := sun, PT := shade_delay);

	IF UP AND DN AND enable AND sun_delay.Q AND cx.SUN_HOR > direction - angle_offset AND cx.SUN_HOR < direction + angle_offset AND
		DT_TO_TOD2(cx.UTC) > cx.SUN_RISE + TIME_TO_UDINT2(sunrise_offset) AND DT_TO_TOD2(cx.UTC) < cx.SUN_SET - TIME_TO_UDINT2(sunset_preset) THEN
		status := BYTE#151;
		QU := UP;
		QD := DN;
		po := shade_pos;
		angle := DEG(ATAN(slat_spacing / slat_width));
		IF cx.SUN_VER > 0.0 AND cx.SUN_VER < angle THEN
			angle := cx.SUN_VER + DEG(ACOS(COS(RAD(cx.SUN_VER))*slat_spacing / Slat_width));
			ao := INT_TO_BYTE(LIMIT(0,UDINT_TO_INT(TRUNC_UDINT2(angle * 2.833333333)), 255));
		ELSE
			ao := BYTE#255;
		END_IF;
	ELSE
		QU := UP;
		QD := DN;
		po := pi;
		ao := ai;
		status := S_IN;
	END_IF;

END_FUNCTION_BLOCK

PROGRAM program0
	VAR
		UP :	BOOL;
		DN :	BOOL;
		S_IN :	BYTE;
		PI :	BYTE;
		AI :	BYTE;
		ENABLE :	BOOL;
		SUN :	BOOL;
		SUNRISE_OFFSET :	TIME := T#1h;
		SUNSET_PRESET :	TIME := T#1h;
		DIRECTION :	REAL := 180.0;
		ANGLE_OFFSET :	REAL := 80.0;
		SLAT_WIDTH :	REAL := 80.0;
		SLAT_SPACING :	REAL := 60.0;
		SHADE_DELAY :	TIME := T#60s;
		SHADE_POS :	BYTE;
		CX :	oscat_CALENDAR;

		func_block : BLIND_SHADE_Block;
	END_VAR
	func_block.UP := UP;
	func_block.DN := DN;
	func_block.S_IN := S_IN ;
	func_block.PI    := PI    ;
	func_block.AI    := AI    ;
	func_block.ENABLE := ENABLE;
	func_block.SUN := SUN;
	func_block.SUNRISE_OFFSET := SUNRISE_OFFSET;
	func_block.SUNSET_PRESET := SUNSET_PRESET ;
	func_block.DIRECTION := DIRECTION ;
	func_block.ANGLE_OFFSET    := ANGLE_OFFSET    ;
	func_block.SLAT_WIDTH := SLAT_WIDTH;
	func_block.SLAT_SPACING := SLAT_SPACING;
	func_block.SHADE_DELAY := SHADE_DELAY ;
	func_block.CX := CX ;

	func_block();
	CX  := func_block.CX;
END_PROGRAM

CONFIGURATION Config0
	RESOURCE Res0 ON PLC
		TASK task0(INTERVAL := T#20ms,PRIORITY := 0);
		PROGRAM instance0 WITH task0 : program0;
	END_RESOURCE
END_CONFIGURATION

(* ---- BLIND_SHADE_S.ST ---- *)
TYPE
  oscat_STRING5               : STRING;
  oscat_STRING30              : STRING;
END_TYPE

TYPE oscat_CALENDAR :
	STRUCT
		UTC : UDINT;				(* world time UTC *)
		LDT : UDINT;				(* local time *)
		LDATE : UDINT;				(* local date *)
		LTOD : UDINT;				(* local time of day *)
		YEAR : INT;					(* year of LDATE *)
		MONTH : INT;				(* month of LDATE *)
		DAY : INT;					(* day of LDATE *)
		WEEKDAY : INT;				(* weekday of LDATE *)
		OFFSET : INT;				(* Time Zone Offset for Local time in minutes *)
		DST_EN : BOOL;				(* daylight savings time enable *)
		DST_ON : BOOL;				(* true when daylight savings time os on *)
		NAME : oscat_string5;		(* name of time zone *)
		LANGUAGE : INT;			    (* language number pls see language setup *)
		LONGITUDE : REAL;			(* longitude of current location *)
		LATITUDE : REAL;			(* latitude of current location *)
		SUN_RISE : UDINT;			(* sun_rise for current location *)
		SUN_SET : UDINT;			(* sun_set for current location *)
		SUN_MIDDAY : UDINT;			(* worldtime when sun stands at south position *)
		SUN_HEIGTH : REAL;			(* suns heigth at midday, south position *)
		SUN_HOR : REAL;				(* sun angle horizontal 0 = north in degrees *)
		SUN_VER : REAL;				(* sun angle vertical above horizon in degrees *)
		NIGHT : BOOL;				(* true between sun_set and sun_rise *)
		HOLIDAY : BOOL;				(* true when holiday *)
		HOLY_NAME : oscat_string30;	(* name of holiday *)
		WORK_WEEK : INT;			(* current work week *)
	END_STRUCT;
END_TYPE

FUNCTION DT_TO_TOD2:UDINT
	VAR_INPUT
		IN :	UDINT;
	END_VAR

	DT_TO_TOD2 := (IN MOD UDINT#86400) * UDINT#1000;
END_FUNCTION

FUNCTION TIME_TO_UDINT2:UDINT
	VAR_INPUT
		X :	TIME;
	END_VAR

	TIME_TO_UDINT2 := DINT_TO_UDINT(TIME_TO_DINT(X));
END_FUNCTION

FUNCTION_BLOCK BLIND_SHADE_S_Block

	VAR_INPUT
		UP :	BOOL;
		DN :	BOOL;
		S_IN :	BYTE;
		PI :	BYTE;
		ENABLE :	BOOL;
		SUN :	BOOL;
		HORZ1 :	REAL := 100.0;
		HORZ2 :	REAL := 260.0;
		VERT :	REAL := 90.0;
		ALERT :	BOOL;
		SUNRISE_OFFSET :	TIME := T#1h;
		SUNSET_PRESET :	TIME := T#1h;
		SHADE_DELAY :	TIME := T#60s;
		SHADE_POS :	BYTE;
		QU :	BOOL;
		QD :	BOOL;
		STATUS :	BYTE;
		PO :	BYTE;
	END_VAR

	VAR_IN_OUT
		CX :	oscat_CALENDAR;
	END_VAR

	VAR
		angle :	REAL;
		sun_delay :	TOF;
	END_VAR

	sun_delay(IN := sun, PT := shade_delay);

	IF ALERT THEN
	QU := TRUE;
	QD := FALSE;
	STATUS := BYTE#152;
	ELSIF UP AND DN AND ENABLE AND sun_delay.Q
	AND (CX.SUN_HOR > HORZ1) AND (CX.SUN_HOR < HORZ2)
	AND (CX.SUN_VER < VERT)
	AND (DT_TO_TOD2(CX.UTC) > CX.SUN_RISE + TIME_TO_UDINT2(sunrise_offset)) AND (DT_TO_TOD2(CX.UTC) < CX.SUN_SET - TIME_TO_UDINT2(sunset_preset)) THEN
	QU := UP;
	QD := DN;
	STATUS := BYTE#151;
	PO := MIN(PI, shade_pos);
	ELSE
	QU := UP;
	QD := DN;
	PO := PI;
	STATUS := S_IN;
	END_IF;

END_FUNCTION_BLOCK

PROGRAM program0
	VAR
		UP :	BOOL;
		DN :	BOOL;
		S_IN :	BYTE;
		PI :	BYTE;
		ENABLE :	BOOL;
		SUN :	BOOL;
		HORZ1 :	REAL := 100.0;
		HORZ2 :	REAL := 260.0;
		VERT :	REAL := 90.0;
		ALERT :	BOOL;
		SUNRISE_OFFSET :	TIME := T#1h;
		SUNSET_PRESET :	TIME := T#1h;
		SHADE_DELAY :	TIME := T#60s;
		SHADE_POS :	BYTE;
		QU :	BOOL;
		QD :	BOOL;
		STATUS :	BYTE;
		PO :	BYTE;
		CX :	oscat_CALENDAR;

		func_block : BLIND_SHADE_S_Block;
	END_VAR
	func_block.UP := UP;
	func_block.DN := DN;
	func_block.S_IN := S_IN ;
	func_block.PI    := PI    ;
	func_block.ENABLE := ENABLE;
	func_block.SUN := SUN;
	func_block.HORZ1 := HORZ1 ;
	func_block.HORZ2 := HORZ2 ;
	func_block.VERT    := VERT    ;
	func_block.ALERT := ALERT;
	func_block.SUNRISE_OFFSET := SUNRISE_OFFSET;
	func_block.SUNSET_PRESET := SUNSET_PRESET ;
	func_block.SHADE_DELAY := SHADE_DELAY ;
	func_block.SHADE_POS    := SHADE_POS    ;
	func_block.QU := QU;
	func_block.QD := QD;
	func_block.STATUS := STATUS ;
	func_block.PO := PO ;
	func_block.CX := CX ;

	func_block();
	CX  := func_block.CX;
END_PROGRAM

CONFIGURATION Config0
	RESOURCE Res0 ON PLC
		TASK task0(INTERVAL := T#20ms,PRIORITY := 0);
		PROGRAM instance0 WITH task0 : program0;
	END_RESOURCE
END_CONFIGURATION

(* ---- BOILER.ST ---- *)
FUNCTION_BLOCK BOILER_Block

	VAR_INPUT
		T_UPPER :	REAL;
		T_LOWER :	REAL;
		PRESSURE :	BOOL := TRUE;
		ENABLE :	BOOL := TRUE;
		REQ_1 :	BOOL;
		REQ_2 :	BOOL;
		BOOST :	BOOL;
		T_UPPER_MIN :	REAL := REAL#50.0;
		T_UPPER_MAX :	REAL := REAL#60.0;
		T_LOWER_ENABLE :	BOOL;
		T_LOWER_MAX :	REAL := REAL#60.0;
		T_REQUEST_1 :	REAL := REAL#70.0;
		T_REQUEST_2 :	REAL := REAL#50.0;
		T_REQUEST_HYS :	REAL := REAL#5.0;
		T_PROTECT_HIGH :	REAL := REAL#80.0;
		T_PROTECT_LOW :	REAL := REAL#10.0;
	END_VAR

	VAR_OUTPUT
		HEAT :	BOOL;
		ERROR :	BOOL;
		STATUS :	BYTE;
	END_VAR

	VAR
		edge :	BOOL;
		boost_mode :	BOOL;
		flag_0 :	BOOL;
		flag_1 :	BOOL;
		flag_2 :	BOOL;
	END_VAR

	IF t_upper > t_protect_high THEN
		status := BYTE#1;
		heat := FALSE;
		error := TRUE;
	ELSIF t_upper < t_protect_low THEN
		status := BYTE#2;
		heat := TRUE;
		error := TRUE;
	ELSIF t_lower > T_protect_high AND t_lower_enable THEN
		status := BYTE#3;
		heat := FALSE;
		error := TRUE;
	ELSIF t_lower < t_protect_low AND t_lower_enable THEN
		status := BYTE#4;
		heat := TRUE;
		error := TRUE;
	ELSIF NOT pressure THEN
		status := BYTE#5;
		heat := FALSE;
		error := TRUE;
	ELSIF req_1 OR req_2 OR enable OR boost THEN
		error := FALSE;

		IF boost AND NOT edge AND t_upper < t_upper_max THEN
			status := BYTE#101;
			heat := TRUE;
			boost_mode := TRUE;
		ELSIF enable AND t_upper < T_upper_min THEN
			status := BYTE#102;
			heat := TRUE;
		ELSIF req_1 AND t_upper < T_request_1 THEN
			status := BYTE#103;
			heat := TRUE;
		ELSIF req_2 AND t_upper < t_request_2 THEN
			status := BYTE#104;
			heat := TRUE;
		END_IF;

		IF heat THEN
			IF (enable OR boost_mode) THEN
				flag_0 := TRUE;
				IF T_lower_enable AND T_lower > T_lower_max THEN
					flag_0 := FALSE;
					boost_mode := FALSE;
				ELSIF NOT T_lower_enable AND T_upper > T_upper_max THEN
					flag_0 := FALSE;
					boost_mode := FALSE;
				END_IF;
			ELSE
				flag_0 := FALSE;
			END_IF;
			flag_1 := (req_1 AND T_upper > T_request_1 + T_request_hys) AND req_1;
			flag_2 := (req_2 AND T_upper > T_request_2 + T_request_hys) AND req_2;

			heat := flag_0 OR flag_1 OR flag_2;
			IF heat = FALSE THEN status := BYTE#100; END_IF;
		END_IF;
	ELSE
		status := BYTE#100;
		heat := FALSE;
		error := FALSE;
	END_IF;
	edge := boost;

END_FUNCTION_BLOCK

PROGRAM program0
	VAR
		T_UPPER :	REAL;
		T_LOWER :	REAL;
		PRESSURE :	BOOL := TRUE;
		ENABLE :	BOOL := TRUE;
		REQ_1 :	BOOL;
		REQ_2 :	BOOL;
		BOOST :	BOOL;
		T_UPPER_MIN :	REAL := REAL#50.0;
		T_UPPER_MAX :	REAL := REAL#60.0;
		T_LOWER_ENABLE :	BOOL;
		T_LOWER_MAX :	REAL := REAL#60.0;
		T_REQUEST_1 :	REAL := REAL#70.0;
		T_REQUEST_2 :	REAL := REAL#50.0;
		T_REQUEST_HYS :	REAL := REAL#5.0;
		T_PROTECT_HIGH :	REAL := REAL#80.0;
		T_PROTECT_LOW :	REAL := REAL#10.0;
		HEAT :	BOOL;
		ERROR :	BOOL;
		STATUS :	BYTE;

		func_block : BOILER_Block;
	END_VAR
	func_block.T_UPPER := T_UPPER;
	func_block.T_LOWER := T_LOWER;
	func_block.PRESSURE := PRESSURE ;
	func_block.ENABLE    := ENABLE    ;
	func_block.REQ_1 := REQ_1;
	func_block.REQ_2 := REQ_2;
	func_block.BOOST := BOOST ;
	func_block.T_UPPER_MIN := T_UPPER_MIN ;
	func_block.T_UPPER_MAX    := T_UPPER_MAX    ;
	func_block.T_LOWER_ENABLE := T_LOWER_ENABLE;
	func_block.T_LOWER_MAX := T_LOWER_MAX;
	func_block.T_REQUEST_1 := T_REQUEST_1 ;
	func_block.T_REQUEST_2 := T_REQUEST_2 ;
	func_block.T_REQUEST_HYS    := T_REQUEST_HYS    ;
	func_block.T_PROTECT_HIGH := T_PROTECT_HIGH;
	func_block.T_PROTECT_LOW := T_PROTECT_LOW;

	func_block();
	HEAT  := func_block.HEAT;
	ERROR  := func_block.ERROR;
	STATUS  := func_block.STATUS;
END_PROGRAM

CONFIGURATION Config0
	RESOURCE Res0 ON PLC
		TASK task0(INTERVAL := T#20ms,PRIORITY := 0);
		PROGRAM instance0 WITH task0 : program0;
	END_RESOURCE
END_CONFIGURATION

(* ---- BOOL_TO_STRING.ST ---- *)
TYPE
  oscat_STRING1               : STRING(1);
END_TYPE

FUNCTION_BLOCK BOOL_TO_STRING_Block
	VAR_INPUT
		IN :	BOOL;
	END_VAR

	VAR_OUTPUT
		BOOL_TO_STRING :	oscat_STRING1;
	END_VAR

	BOOL_TO_STRING := SEL_STRING(IN,'0','1');
END_FUNCTION_BLOCK

PROGRAM program0
  VAR
    LocalVar0 : BOOL;
	LocalOUT  : oscat_STRING1;
	func_block : BOOL_TO_STRING_Block;
  END_VAR
	func_block.IN := LocalVar0;
	func_block();
	LocalOUT := func_block.BOOL_TO_STRING;

END_PROGRAM

CONFIGURATION Config0
  RESOURCE Res0 ON PLC
    TASK task0(INTERVAL := T#20ms,PRIORITY := 0);
    PROGRAM instance0 WITH task0 : program0;
  END_RESOURCE
END_CONFIGURATION

(* ---- BUFFER_CLEAR.ST ---- *)
TYPE
	oscat_arb_0_249 			  : ARRAY [0..249] 	OF BYTE;
END_TYPE

FUNCTION_BLOCK _BUFFER_CLEAR
	VAR_IN_OUT
		PT :	oscat_arb_0_249;
	END_VAR

	VAR_INPUT
		SIZE :	UINT;
	END_VAR

	VAR_OUTPUT
		BUFFER_CLEAR :	BOOL;
	END_VAR

	VAR
		err :	INT;
		result :	WORD;
	END_VAR

	result := MEMSET(err,BYTE#00,UINT_TO_DINT(size),pt[0]);
	BUFFER_CLEAR := (err = 0);

END_FUNCTION_BLOCK

PROGRAM program0
	VAR
	    LocalVar1 : oscat_arb_0_249;
		LocalVar2 : UINT;
		LocalOUT  : BOOL;
		func_block : _BUFFER_CLEAR;
  	END_VAR
	func_block.PT := LocalVar1;
	func_block.SIZE := LocalVar2;
	func_block();
	LocalOUT := func_block.BUFFER_CLEAR;
END_PROGRAM

CONFIGURATION Config0
	VAR_GLOBAL
		PLC_TICKS_PER_SEC :	INT;
		PLC_SYS_TICK_CNT :	DINT;
	END_VAR

  	RESOURCE Res0 ON PLC
    	TASK task0(INTERVAL := T#20ms,PRIORITY := 0);
    	PROGRAM instance0 WITH task0 : program0;
  	END_RESOURCE
END_CONFIGURATION

(* ---- BUFFER_CLEAR_NW.ST ---- *)
TYPE
  oscat_NW_BUF_LONG  : ARRAY [0..4095] OF BYTE;
END_TYPE

FUNCTION_BLOCK _BUFFER_CLEAR_NW
	VAR_INPUT
		SIZE :	UINT;
	END_VAR

	VAR_OUTPUT
		BUFFER_CLEAR :	BOOL;
	END_VAR

	VAR_IN_OUT
		PT :	oscat_NW_BUF_LONG;
	END_VAR

	VAR
		err :	INT;
		result :	WORD;
	END_VAR
	result:=MEMSET(err,BYTE#00,UINT_TO_DINT(size),pt[0]);
	BUFFER_CLEAR := (err = 0);
END_FUNCTION_BLOCK

PROGRAM program0
  VAR
	SIZE :	UINT;

	BUFFER_CLEAR :	BOOL;

	PT :	oscat_NW_BUF_LONG;

	func_block : _BUFFER_CLEAR_NW;
  END_VAR
	func_block.SIZE  :=SIZE ;
	func_block.PT  :=PT ;
	func_block();
	PT := func_block.PT;
	BUFFER_CLEAR := func_block.BUFFER_CLEAR;
END_PROGRAM

CONFIGURATION Config0
  RESOURCE Res0 ON PLC
    TASK task0(INTERVAL := T#20ms,PRIORITY := 0);
    PROGRAM instance0 WITH task0 : program0;
  END_RESOURCE
END_CONFIGURATION

(* ---- BUFFER_COMP.ST ---- *)
TYPE
	oscat_arb_0_249 			  : ARRAY [0..249] 	OF BYTE;
END_TYPE

FUNCTION_BLOCK BUFFER_COMP_Block
	VAR_IN_OUT
		PT1 :	oscat_arb_0_249;
	END_VAR

	VAR_INPUT
		SIZE1 :	INT;
	END_VAR

	VAR_IN_OUT
		PT2 :	oscat_arb_0_249;
	END_VAR

	VAR_INPUT
		SIZE2 :	INT;
		START :	INT;
	END_VAR

	VAR_OUTPUT
		BUFFER_COMP :	INT;
	END_VAR

	VAR
		i :	INT;
		j :	INT;
		end :	INT;
		j2 :	INT;
	END_VAR

	IF SIZE2 <= SIZE1 AND SIZE1 > 0 AND SIZE2 > 0 AND START >= 0 THEN
		end := SIZE1 - SIZE2;
		FOR i := START TO end DO
			IF PT1[i] = PT2[0] THEN
				(* first character matches, now compare rest of array *)
				j := 1;
				j2 := j + i;
				WHILE j < SIZE2 DO
					IF PT2[j] <> PT1[j2] THEN EXIT; END_IF;
					j := j + 1;
					j2 := j2 + 1;
				END_WHILE;
				(* when J > size2 a match was found return the position i in buffer1 *)
				IF j = SIZE2 THEN
					BUFFER_COMP := i;
					RETURN;
				END_IF;
			END_IF;
		END_FOR;
	END_IF;
	BUFFER_COMP := -1;

END_FUNCTION_BLOCK

PROGRAM program0
  VAR
    LocalVar0 : oscat_arb_0_249;
    LocalVar1 : INT;
	LocalVar2 : oscat_arb_0_249;
	LocalVar3 : INT;
	LocalVar4 : INT;
	LocalOUT  : INT;
	func_block : BUFFER_COMP_Block;
  END_VAR
	func_block.PT1  := LocalVar0;
	func_block.SIZE1 := LocalVar1;
	func_block.PT2  := LocalVar2;
	func_block.SIZE2 := LocalVar3;
	func_block.START := LocalVar4;
	func_block();
	LocalOUT := func_block.BUFFER_COMP;
	LocalVar0 := func_block.PT1;
	LocalVar2 := func_block.PT1;

END_PROGRAM

CONFIGURATION Config0
  RESOURCE Res0 ON PLC
    TASK task0(INTERVAL := T#20ms,PRIORITY := 0);
    PROGRAM instance0 WITH task0 : program0;
  END_RESOURCE
END_CONFIGURATION

(* ---- BUFFER_COMP_NW.ST ---- *)
TYPE
  oscat_NW_BUF_LONG  : ARRAY [0..4095] OF BYTE;
END_TYPE

FUNCTION_BLOCK BUFFER_COMP_NW
	VAR_IN_OUT
		PT1 :	oscat_NW_BUF_LONG;
	END_VAR

	VAR_INPUT
		SIZE1 :	INT;
	END_VAR

	VAR_IN_OUT
		PT2 :	oscat_NW_BUF_LONG;
	END_VAR

	VAR_INPUT
		SIZE2 :	INT;
		START :	INT;
	END_VAR

	VAR_OUTPUT
		BUFFER_COMP :	INT;
	END_VAR

	VAR
		i :	INT;
		j :	INT;
		end :	INT;
		j2 :	INT;
	END_VAR

	IF SIZE2 <= SIZE1 AND SIZE1 > 0 AND SIZE2 > 0 AND START >= 0 THEN
		end := SIZE1 - SIZE2;
		FOR i := START TO end DO
			IF PT1[i] = PT2[0] THEN
				(* first character matches, now compare rest of array *)
				j := 1;
				j2 := j + i;
				WHILE j < SIZE2 DO
					IF PT2[j] <> PT1[j2] THEN EXIT; END_IF;
					j := j + 1;
					j2 := j2 + 1;
				END_WHILE;
				(* when J > size2 a match was found return the position i in buffer1 *)
				IF j = SIZE2 THEN
					BUFFER_COMP := i;
					RETURN;
				END_IF;
			END_IF;
		END_FOR;
	END_IF;
	BUFFER_COMP := -1;

END_FUNCTION_BLOCK

PROGRAM program0
  VAR
	PT1   :	oscat_NW_BUF_LONG;

	SIZE1 :	INT;

	PT2   : 	oscat_NW_BUF_LONG;

	SIZE2 :	INT;
	START :	INT;

	BUFFER_COMP :	INT;

	func_block : BUFFER_COMP_NW;
  END_VAR
	func_block.PT1  :=PT1  ;
	func_block.SIZE1:=SIZE1;
	func_block.PT2  :=PT2  ;
	func_block.SIZE2:=SIZE2;
	func_block.START:=START;
	func_block();
	BUFFER_COMP := func_block.BUFFER_COMP;
	PT1 := func_block.PT1;
	PT2 := func_block.PT2;

END_PROGRAM

CONFIGURATION Config0
  RESOURCE Res0 ON PLC
    TASK task0(INTERVAL := T#20ms,PRIORITY := 0);
    PROGRAM instance0 WITH task0 : program0;
  END_RESOURCE
END_CONFIGURATION

(* ---- BUFFER_INSERT_NW.ST ---- *)
TYPE
  oscat_NW_BUF_LONG  : ARRAY [0..4095] OF BYTE;
END_TYPE

FUNCTION_BLOCK _BUFFER_INSERT_NW
	VAR_INPUT
		STR :	STRING;
		POS :	INT;
	END_VAR

	VAR_IN_OUT
		PT :	oscat_NW_BUF_LONG;
	END_VAR

	VAR_INPUT
		SIZE :	UINT;
	END_VAR

	VAR_OUTPUT
		_BUFFER_INSERT :	INT;
	END_VAR

	VAR
		end :	INT;
		lx :	INT;
		i :	INT;
		i2 :	INT;
		_STRING_TO_BUFFER :	_STRING_TO_BUFFER;
	END_VAR

	i := UINT_TO_INT(size) - 1;
	pos := LIMIT_INT(0,pos,i);
	lx := LEN(str);
	end := pos + lx;
	(* first move the upper part of the buffer to make space for the string *)
	i2 := i - lx;
	WHILE i >= end DO
	pt[i] := pt[i2];
	i  := i  - 1;
	i2 := i2 - 1;
	END_WHILE;

	_STRING_TO_BUFFER(str:=str, pos:=pos, size:=size, pt:=pt);
	_BUFFER_INSERT := _STRING_TO_BUFFER._STRING_TO_BUFFER;
	pt := _STRING_TO_BUFFER.pt;
END_FUNCTION_BLOCK

PROGRAM program0
  VAR
	STR :	STRING;
	POS :	INT;

	PT :	oscat_NW_BUF_LONG;

	SIZE :	UINT;

	_BUFFER_INSERT :	INT;
	func_block : _BUFFER_INSERT_NW;
  END_VAR
	func_block.STR  :=STR ;
	func_block.POS  :=POS ;
	func_block.SIZE  :=SIZE ;
	func_block.PT  :=PT ;
	func_block();
	PT := func_block.PT;
	_BUFFER_INSERT := func_block._BUFFER_INSERT;
END_PROGRAM

CONFIGURATION Config0
  RESOURCE Res0 ON PLC
    TASK task0(INTERVAL := T#20ms,PRIORITY := 0);
    PROGRAM instance0 WITH task0 : program0;
  END_RESOURCE
END_CONFIGURATION

(* ---- BUFFER_SEARCH.ST ---- *)
TYPE
	oscat_arb_0_249 			  : ARRAY [0..249] 	OF BYTE;
END_TYPE

FUNCTION_BLOCK BUFFER_SEARCH_Block
	VAR_INPUT
		SIZE :	UINT;
		STR :	STRING;
		POS :	INT;
		IGN :	BOOL;
	END_VAR

	VAR_IN_OUT
		PT :	oscat_arb_0_249;
	END_VAR

	VAR_OUTPUT
		BUFFER_SEARCH :	INT;
	END_VAR

	VAR
		i :	INT;
		end :	INT;
		k :	INT;
		k2 :	INT;
		lx :	INT;
		char :	BYTE;
		chx :	BYTE;
	END_VAR

	lx := LEN(str);
	IF pos >= 0 AND lx > 0 THEN
		end := UINT_TO_INT(size) - lx;
		lx := lx - 1;
		FOR i := pos TO end DO
			FOR k := 0 TO lx DO
				char := INT_TO_BYTE(GET_CHAR(str,k + 1));
				k2 := i + k;
				IF IGN THEN
					chx := TO_UPPER(pt[k2]);
				ELSE
					chx := pt[k2];
				END_IF;
				IF char <> chx THEN EXIT; END_IF;
			END_FOR;
			IF k > lx THEN
				BUFFER_SEARCH := i;
				RETURN;
			END_IF;
		END_FOR;
	END_IF;
	BUFFER_SEARCH := -1;
END_FUNCTION_BLOCK

PROGRAM program0
  VAR
    LocalVar0 : UINT;
    LocalVar1 : STRING;
	LocalVar2 : INT;
	LocalVar3 : BOOL;
	LocalVar4 : oscat_arb_0_249;
	LocalOUT  : INT;
	func_block : BUFFER_COMP_Block;
  END_VAR
	func_block.SIZE  := LocalVar0;
	func_block.STR  := LocalVar1;
	func_block.POS   := LocalVar2;
	func_block.IGN  := LocalVar3;
	func_block.PT := LocalVar4;
	func_block();
	LocalOUT := func_block.BUFFER_COMP;
	LocalVar4 := func_block.PT;

END_PROGRAM

CONFIGURATION Config0
  RESOURCE Res0 ON PLC
    TASK task0(INTERVAL := T#20ms,PRIORITY := 0);
    PROGRAM instance0 WITH task0 : program0;
  END_RESOURCE
END_CONFIGURATION

(* ---- BUFFER_TO_STRING.ST ---- *)
TYPE
	oscat_arb_0_249 			  : ARRAY [0..249] 	OF BYTE;
END_TYPE

FUNCTION_BLOCK BUFFER_TO_STRING_Block
	VAR_IN_OUT
		PT  :	oscat_arb_0_249;
	END_VAR

	VAR_INPUT
		SIZE :	UINT;
		START :	UINT;
		STOP :	UINT;
	END_VAR

	VAR_OUTPUT
		BUFFER_TO_STRING :	STRING;
	END_VAR

	VAR
		sta :	UINT;
		stp :	UINT;
		size2 :	UINT;
		i :	INT;
		BUF_TO_STRING :	BUF_TO_STRING;
	END_VAR

	sta := MIN(START, SIZE - UINT#1);
	stp := STOP;
	IF stp - sta + UINT#1 > UINT#250 THEN
		stp := sta + UINT#250 - UINT#1;
	END_IF;
	stp := MIN(stp, SIZE - UINT#1);
	size2 := stp - sta + UINT#1;
	IF size2 > UINT#0 THEN
		FOR i := 0 TO 1 DO
			BUF_TO_STRING.REQ := i > 0;
			BUF_TO_STRING.BUF_FORMAT := TRUE;
			BUF_TO_STRING.BUF_OFFS := UINT_TO_DINT(START);
			BUF_TO_STRING.BUF_CNT := UINT_TO_DINT(size2);
			BUF_TO_STRING.BUFFER := pt;
			BUF_TO_STRING.DST := BUFFER_TO_STRING;
			BUF_TO_STRING();
			pt := BUF_TO_STRING.BUFFER;
			BUFFER_TO_STRING := BUF_TO_STRING.DST;
		END_FOR;
	ELSE
		BUFFER_TO_STRING :='';
	END_IF;
END_FUNCTION_BLOCK

PROGRAM program0
  VAR
    LocalVar0 : oscat_arb_0_249;
    LocalVar1 : UINT;
	LocalVar2 : UINT;
	LocalVar3 : UINT;
	LocalOUT  : INT;
	func_block : BUFFER_TO_STRING_Block;
  END_VAR
	func_block.PT  := LocalVar0;
	func_block.SIZE := LocalVar1;
	func_block.START := LocalVar2;
	func_block.STOP := LocalVar3;
	func_block();
	LocalOUT := func_block.BUFFER_TO_STRING;
	LocalVar0 := func_block.PT;

END_PROGRAM

CONFIGURATION Config0
  RESOURCE Res0 ON PLC
    TASK task0(INTERVAL := T#20ms,PRIORITY := 0);
    PROGRAM instance0 WITH task0 : program0;
  END_RESOURCE
END_CONFIGURATION
